(* IEC 61131-3 sources: daoli-st-library/DL_Device (part 29) *)

(* ---- FB_DL_PulseFlowMeter.st ---- *)
(*==============================================================================
 * 组件名称 (Component)  : FB_DL_PulseFlowMeter
 * 所属子库 (Sublibrary) : DL_Device
 * 当前版本 (Version)    : 1.0.0
 * 兼容性   (Platform)   : CODESYS 3.5 / TwinCAT 3 / 汇川 InoProShop / Machine Expert
 *                         仅依赖 Standard.library（TON / R_TRIG），零厂商方言
 * 分类     (Category)   : 设备功能块（Function Block，实现 I_DL_FlowMeter）
 * 功能简述 (Function)   : 脉冲型流量计瞬时流量与累计总量计量。脉冲沿计数 →
 *                         自重触发采样窗频率估计 → K 系数换算 [L/min]；总量
 *                         按脉冲计数法累计（精度优于流量积分法）；低流量截
 *                         止、脉冲丢失超时、频率超量程提示；K 系数防除零。
 *                         滑动窗计数为 Device 层内联实现（依赖方向合规：不
 *                         引 DL_MathData 组件）。
 * 接口实现 (Implements) : I_DL_FlowMeter。接口属性同名成员（eState/fFlowRate/
 *                         fTotal/nPulseCount/bFault/uErrorId）按 R22 以只读
 *                         PROPERTY GET 承载（内部镜像同源），非接口成员
 *                         bTotalNearLimit 保留 VAR_OUTPUT；方法 CmdTotalReset/
 *                         CmdTotalPreset/CmdReset 在本文件尾部落地。
 * 公约遵循 (Convention) : 0.1/R23 周期计量型（无初始化/跟踪同步语义，窗由自
 *                         重触发 TON 驱动），免首扫，无 bInit。
 *                         0.2/R21 bFault 显式排除信息级码；0.5/R7 全部实例主
 *                         体最前部无条件刷新；0.7/R15 故障级锁存仅复位路径清
 *                         码；0.9 全部 REAL/LREAL 输入先做非数自比检测再比
 *                         较，出口默认值在第一条防御 IF 之前赋值。
 *                         0.8 故障码段位 16#0003_xxxx（经 DL_Device
 *                         VERSION.md 码表核对：规格建议信息级 0003_0107/
 *                         0108/0109 已被 FB_DL_VfdGeneric/FB_DL_AnalogValve
 *                         占用，依公约冲突顺延）：
 *                         【故障级】0003_02B0 K 系数非法；
 *                         【信息级】0003_0113 低流量截止激活、0003_0114 脉冲
 *                         丢失超时、0003_0115 窗内频率超量程。
 * 红线自检 (Redline)    : R1 零全局变量表/外部变量引用 ✓｜R2 零物理 IO 地址 ✓
 *                         R3 纯 IEC 61131-3 ✓｜R4 三处除法全部带 ABS(分母)
 *                         >1E-6 防零分支并置码 ✓
 *                         R5 全变量中英双语同行注释 ✓｜R6 状态映像 IF 派生链
 *                         含 ELSE 兜底（无显式 CASE 主状态机，计量型派生映
 *                         像）✓
 *                         R7 四实例（R_TRIG×3/TON×2）主体最前部无条件刷新 ✓
 *                         R8 全常量化 ✓
 * 设计要点 (Key notes)  : ① 瞬时流量 = 窗脉冲数 / 窗秒数 / fKFactor × 60；
 *                         ② 双缓冲：窗运行期脉冲进计数缓冲，窗沿（TON 振荡
 *                           器 Q）整窗交换到读出缓冲，读侧永不撕裂；
 *                         ③ 除零防御三处：fKFactor 非法 → 故障锁存；窗秒数
 *                           由钳位域（100MS~10S）恒非零 + 显式 ABS 防零分支；
 *                           周期法不使用（统一窗法，简化跨平台）；
 *                         ④ 总量按脉冲计数法 fTotal += 窗脉冲数 / fKFactor；
 *                         ⑤ fTotal > 9.0E15 预警（LREAL 整数精度边界）。
 * 偏离留档 (Deviation)  : 依 R11 头注释留档，共 1 条：
 *                         ① 信息级码顺延：规格建议 0003_0107/0108/0109 与既
 *                           有组件冲突，依公约 0.8 顺延为 0003_0113/0114/
 *                           0115（核对结果优先于建议值）。
 * 开源溯源 (Origin)     : 来源标签 tcopen-component / flow-totalizer，T1-1
 *                         OSCAT Basic ◐ 深化旁证（RAW_NOTES_R7 S-6：TcOpen
 *                         流量组件语义域 + OSCAT 流量计窗法计数公开实现思
 *                         想，仅借鉴语义与算法思想；双缓冲、码位与引脚契约
 *                         100% 本库独立设计，clean-room 未复制源码）。
 * 验收向量 (Acceptance) :
 *   V1 已知脉冲序列换算逐拍复算：窗 1S 内 100 脉冲、K=100 → 1.0 L/min；
 *   V2 总量累计与清零：连续 10 窗 @100 脉冲 → fTotal=10.0 L；清零沿 → 0；
 *   V3 低流量截止：fFlowRate < fLowCutoff → 输出置零 + eLowCutoff + 0003_0113；
 *   V4 K 系数非法：fKFactor=0 → 故障锁存 0003_02B0；
 *   V5 脉冲丢失：tPulseTimeout 超时无脉冲 → 流量置零 + 0003_0114；
 *   V6 双缓冲无撕裂推演：窗沿交换拍读侧保持整窗旧值，计数侧从零重启。
 * 修订历史 (Revision)   :
 *   2026-11-15  v1.0.0  首版入库（Round 07 · DL_Device 流量计族实现件）
 *============================================================================*)
FUNCTION_BLOCK FB_DL_PulseFlowMeter IMPLEMENTS I_DL_FlowMeter
VAR_INPUT
    bPulseIn       : BOOL;             // 脉冲输入（Pulse input），R_TRIG 上升沿计数；硬件滤波由输入层保证 / Pulse input, counted on rising edge, HW filtering upstream
    bCmdTotalReset : BOOL;             // 总量清零指令（Total reset command），上升沿生效 / Total reset edge
    fKFactor       : REAL := 100.0;    // 流量计 K 系数（K-factor）[pulses/L]，域 >0，默认 100.0；标定证书值 / K-factor [pulses/L], > 0, calibration value
    tSampleWindow  : TIME := T#1S;     // 频率估计采样窗（Sample window），默认 T#1S，域 100MS~10S 越界钳位；低流量场景增大 / Sample window, clamped 100MS..10S, increase for low flow
    fLowCutoff     : REAL := 0.5;      // 低流量截止阈值（Low-flow cutoff）[L/min]，默认 0.5；低于阈值输出置零 / Low-flow cutoff [L/min], below it the output is zeroed
    tPulseTimeout  : TIME := T#5S;     // 脉冲丢失超时（Pulse timeout），默认 T#5S；运行中窗口超时无脉冲 → 流量置零 + 信息级 / Pulse timeout, no pulse in window zeroes the flow with info
    bReset         : BOOL;             // 上升沿复位故障（Reset edge）/ Rising edge resets fault
END_VAR
VAR_OUTPUT
    bTotalNearLimit : BOOL;            // 总量接近溢出预警（Total near limit），fTotal > 9.0E15 置位（LREAL 整数精度边界）/ Total near LREAL integer-precision boundary
END_VAR
VAR
    _eState        : E_DL_FlowMeterState := E_DL_FlowMeterState.eIdle; // 内部计量状态（Internal metering state），属性只读 / Internal state, read-only via property
    _bFaultLatch   : BOOL;             // 故障锁存标志（Fault latch flag），仅复位路径清除 / Fault latch, cleared only via reset path
    _uErrorIdInt   : UDINT;            // 内部故障级码寄存（Internal fault-level register）/ Internal fault-level register
    _uInfoCode     : UDINT;            // 本拍信息级码（Info code this cycle），瞬时型每拍重算 / Transient info code, recomputed each scan
    _fKFactorEff   : REAL := 100.0;    // 防御后生效 K 系数（Sanitized K-factor）[pulses/L] / Sanitized K-factor
    _fCutoffEff    : REAL := 0.5;      // 防御后生效截止阈值（Sanitized cutoff）[L/min] / Sanitized cutoff
    _tWindowEff    : TIME := T#1S;     // 钳位后生效采样窗（Clamped sample window）/ Clamped sample window
    _nCounting     : UDINT;            // 计数中缓冲（Counting buffer），窗运行期累积 / Counting buffer during the window
    _nLastWin      : UDINT;            // 读出缓冲（Readout buffer），窗沿整窗交换 / Readout buffer swapped at window edge
    _fTotalInt     : LREAL;            // 内部累计总量（Internal totalized volume）[L] / Internal totalized volume [L]
    _fFlowRateInt  : REAL;             // 内部瞬时流量（Internal flow rate）[L/min] / Internal flow rate [L/min]
    _fWinSec       : REAL := 1.0;      // 窗秒数（Window seconds），TIME 显式换算 / Window length in seconds, explicit conversion
    _bHadPulse     : BOOL;             // 曾收到脉冲标志（Ever-pulsed flag），超时判定前提 / Ever-pulsed flag, timeout precondition
    _bPulseLost    : BOOL;             // 脉冲丢失超时激活（Pulse-lost timeout active）/ Pulse-lost timeout active
    _bLowCutoffAct : BOOL;             // 低流量截止激活标志（Low-flow cutoff active flag）/ Low-flow cutoff active flag
    _bPendTotalRst : BOOL;             // 方法总量清零请求（Method total-reset request）/ Method total-reset request
    _bPendPreset   : BOOL;             // 方法总量预置请求（Method total-preset request）/ Method total-preset request
    _fPresetVal    : LREAL;            // 方法预置值（Method preset value）[L] / Method preset value [L]
    _bPendReset    : BOOL;             // 方法复位请求（Method reset request）/ Method reset request
    _fbTrigPulse   : R_TRIG;           // 脉冲上升沿（Pulse rising edge）/ Pulse edge detector
    _fbTrigTotalRst: R_TRIG;           // 引脚总量清零沿（Pin total-reset edge）/ Pin total-reset edge detector
    _fbTrigReset   : R_TRIG;           // 引脚复位沿（Pin reset edge）/ Pin reset edge detector
    _fbTonWindow   : TON;              // 采样窗振荡器（Sample-window oscillator），IN := NOT Q 自重触发 / Sample-window oscillator, self-retriggered
    _fbTonPulseTo  : TON;              // 脉冲丢失超时（Pulse-lost timeout）/ Pulse-lost timeout
END_VAR
VAR CONSTANT
    DL_WIN_MIN     : TIME := T#100MS;  // 采样窗下限（Sample window lower clamp）/ Sample window lower clamp
    DL_WIN_MAX     : TIME := T#10S;    // 采样窗上限（Sample window upper clamp）/ Sample window upper clamp
    DL_PULSE_WIN_MAX : UDINT := 10000; // 单窗脉冲数超量程阈值（Pulses-per-window overrange limit），提示配置 HSC / Per-window pulse overrange, suggests HSC
    DL_TOTAL_LIMIT : LREAL := 9.0E15;  // 总量精度边界预警阈值（Total precision-boundary threshold）[L] / Total precision-boundary threshold [L]
    DL_REAL_EPS    : REAL := 1.0E-6;   // 浮点防零容差（Float divide-guard epsilon）/ Float divide-guard epsilon
END_VAR

METHOD CmdTotalReset : BOOL
VAR_INPUT
END_VAR
IF _bFaultLatch OR (_eState = E_DL_FlowMeterState.eFault) THEN
    CmdTotalReset := FALSE;       // 故障态拒绝（Rejected in fault）
ELSE
    _bPendTotalRst := TRUE;       // 登记清零请求，主体消化（Register reset, consumed by body）
    CmdTotalReset := TRUE;        // 受理成功（Accepted）
END_IF

(*------------------------------------------------------------------------------
 * 方法: CmdTotalPreset —— 总量预置 [L]，非有限值/负值拒绝返回 FALSE。
 *      Method CmdTotalPreset - total preset [L], non-finite or negative rejected.
 *------------------------------------------------------------------------------*)
    END_METHOD

METHOD CmdTotalPreset : BOOL
VAR_INPUT
    fPreset : LREAL; // 预置总量（Preset volume）[L]，域 ≥0 / Preset volume [L], range >= 0
END_VAR
IF _bFaultLatch OR (_eState = E_DL_FlowMeterState.eFault) THEN
    CmdTotalPreset := FALSE;      // 故障态拒绝（Rejected in fault）
ELSIF (fPreset <> fPreset) OR (fPreset < 0.0) THEN
    CmdTotalPreset := FALSE;      // 非数或负值拒绝（Rejected on NaN or negative）
ELSE
    _fPresetVal := fPreset;       // 登记预置值（Register preset value）
    _bPendPreset := TRUE;         // 登记预置请求（Register preset request）
    CmdTotalPreset := TRUE;       // 受理成功（Accepted）
END_IF

(*------------------------------------------------------------------------------
 * 方法: CmdReset —— 复位故障。仅故障态受理（接口方法拒绝语义红线）。
 *      Method CmdReset - reset, accepted only in fault state.
 *------------------------------------------------------------------------------*)
    END_METHOD

METHOD CmdReset : BOOL
VAR_INPUT
END_VAR
IF _bFaultLatch OR (_eState = E_DL_FlowMeterState.eFault) THEN
    _bPendReset := TRUE;          // 登记复位请求（Register reset request）
    CmdReset := TRUE;             // 可复位（Resettable）
ELSE
    CmdReset := FALSE;            // 无故障可复位（Nothing to reset）
END_IF

(*------------------------------------------------------------------------------
 * 属性: eState（GET）—— 当前计量状态只读视图。
 *      Property eState (GET) - read-only metering state view.
 *------------------------------------------------------------------------------*)
    END_METHOD

// ============================================================================
// 段 1｜实例无条件周期刷新（R7/0.5：严禁置于 IF/CASE 分支内）
//      Unconditional per-cycle refresh of all instances (R7/0.5)
// ============================================================================
_fbTrigPulse(CLK    := bPulseIn);
_fbTrigTotalRst(CLK := bCmdTotalReset);
_fbTrigReset(CLK    := bReset);
_fbTonWindow(IN := (NOT _fbTonWindow.Q) AND (NOT _bFaultLatch), PT := _tWindowEff); // 采样窗振荡器（Window oscillator）
_fbTonPulseTo(IN := _bHadPulse AND (NOT _fbTrigPulse.Q) AND (NOT _bFaultLatch), PT := tPulseTimeout); // 脉冲丢失超时（Pulse-lost timeout）

// ============================================================================
// 段 2｜参数防御（0.9：非数自比检测，出口默认值先行）+ 信息级预清零 + 复位
//      Parameter sanitation (0.9) + info preset + reset path
// ============================================================================
_uInfoCode := 0;                  // 信息级瞬时型每拍重算（Transient info recomputed each scan）

IF fKFactor <> fKFactor THEN      // K 系数非数自比检测（K-factor NaN self-compare）
    _bFaultLatch := TRUE;         // K 系数非法锁存（Invalid K-factor latch）
    _uErrorIdInt := 16#0003_02B0; // 0003_02B0 K 系数非法【故障级】/ Invalid K-factor, fault level
ELSIF ABS(fKFactor) <= DL_REAL_EPS THEN
    _bFaultLatch := TRUE;         // K 系数趋零防除零锁存（Near-zero K-factor latch）
    _uErrorIdInt := 16#0003_02B0; // 0003_02B0 K 系数非法【故障级】/ Invalid K-factor, fault level
ELSE
    _fKFactorEff := fKFactor;     // 生效 K 系数镜像（Effective K-factor mirror）
END_IF

IF fLowCutoff <> fLowCutoff THEN  // 截止阈值非数自比（Cutoff NaN self-compare）
    _fCutoffEff := 0.5;           // 回落默认阈值（Fallback default cutoff）
ELSIF fLowCutoff < 0.0 THEN
    _fCutoffEff := 0.0;           // 负值钳零（Negative clamped to zero）
ELSE
    _fCutoffEff := fLowCutoff;    // 生效阈值镜像（Effective cutoff mirror）
END_IF

IF tSampleWindow < DL_WIN_MIN THEN
    _tWindowEff := DL_WIN_MIN;    // 采样窗下限钳位（Window lower clamp）
ELSIF tSampleWindow > DL_WIN_MAX THEN
    _tWindowEff := DL_WIN_MAX;    // 采样窗上限钳位（Window upper clamp）
ELSE
    _tWindowEff := tSampleWindow; // 合法直通（Valid pass-through）
END_IF
_fWinSec := TIME_TO_REAL(_tWindowEff) / 1000.0; // TIME→REAL 换算结果为毫秒数，除 1000 得秒（CODESYS/TwinCAT 口径，舍入意图：整毫秒窗恒精确）/ TIME_TO_REAL yields milliseconds, divide by 1000 for seconds

IF _fbTrigReset.Q OR _bPendReset THEN
    _bPendReset := FALSE;         // 消费方法复位请求（Consume method reset）
    _bFaultLatch := FALSE;        // 故障锁存解除（Fault latch released）
    _uErrorIdInt := 16#0000_0000; // 故障码清零（Fault code cleared）
END_IF

// ============================================================================
// 段 3｜总量清零/预置（引脚沿 + 方法请求）
//      Total reset/preset (pin edge + method request)
// ============================================================================
IF _fbTrigTotalRst.Q OR _bPendTotalRst THEN
    _bPendTotalRst := FALSE;      // 消费方法请求（Consume method request）
    _fTotalInt := 0.0;            // 总量清零（Total cleared）
END_IF
IF _bPendPreset THEN
    _bPendPreset := FALSE;        // 消费方法预置请求（Consume method preset）
    IF _fPresetVal >= 0.0 THEN
        _fTotalInt := _fPresetVal; // 合法预置写入（Valid preset written）
    END_IF                         // 非法预置已被方法拒绝，此处仅兜底（Invalid preset already rejected by method）
END_IF

// ============================================================================
// 段 4｜脉冲计数 + 窗沿双缓冲交换 + 瞬时流量换算（除法全部带防零分支）
//      Pulse counting + double-buffer swap at window edge + flow conversion
// ============================================================================
IF _fbTrigPulse.Q THEN
    _nCounting := _nCounting + 1; // 计数缓冲累加（Counting buffer increment）
    _bHadPulse := TRUE;           // 曾收到脉冲（Ever pulsed）
END_IF

IF _fbTonWindow.Q THEN
    // 窗沿：整窗交换（双缓冲无撕裂：读出缓冲只在窗沿被写一次）
    // Window edge: whole-window swap (readout written once per window, no tearing)
    _nLastWin := _nCounting;      // 读出缓冲接收整窗计数（Readout takes the window count）
    _nCounting := 0;              // 计数缓冲清零重启（Counting buffer restarted）
    IF ABS(_fKFactorEff) > DL_REAL_EPS THEN
        _fTotalInt := _fTotalInt + UDINT_TO_LREAL(_nLastWin) / _fKFactorEff; // 脉冲计数法累计（Count-based totalization, divisor proven non-zero）
    END_IF
END_IF

_fFlowRateInt := 0.0;             // 出口默认值先赋（Default outlet first）
IF ABS(_fWinSec) > DL_REAL_EPS THEN
    IF ABS(_fKFactorEff) > DL_REAL_EPS THEN
        _fFlowRateInt := UDINT_TO_REAL(_nLastWin) / _fWinSec / _fKFactorEff * 60.0; // 窗法换算 [L/min]（Window-method conversion, divisors proven non-zero）
    END_IF
END_IF

// ============================================================================
// 段 5｜诊断与信息级：脉冲丢失 / 频率超量程 / 低流量截止
//      Diagnostics and info codes: pulse lost / overrange / low-flow cutoff
// ============================================================================
_bLowCutoffAct := FALSE;          // 截止激活标志每拍预清零（Cutoff flag preset FALSE）
_bPulseLost := _fbTonPulseTo.Q;   // 脉冲丢失超时激活（Pulse-lost timeout active）
IF _bPulseLost THEN
    _fFlowRateInt := 0.0;         // 超时流量置零（Flow zeroed on timeout）
    _uInfoCode := 16#0003_0114;   // 0003_0114 脉冲丢失超时【信息级】/ Pulse-lost timeout, info level
ELSIF _nLastWin > DL_PULSE_WIN_MAX THEN
    _uInfoCode := 16#0003_0115;   // 0003_0115 窗内频率超量程【信息级】，提示输入层配置 HSC / Per-window overrange, suggest HSC upstream
ELSIF (_fFlowRateInt < _fCutoffEff) AND _bHadPulse AND (NOT _bPulseLost) THEN
    _fFlowRateInt := 0.0;         // 低流量截止输出置零（Low-flow cutoff zeroes output）
    _bLowCutoffAct := TRUE;       // 截止激活标志置位（Cutoff flag asserted）
    _uInfoCode := 16#0003_0113;   // 0003_0113 低流量截止激活【信息级】/ Low-flow cutoff active, info level
END_IF

// ============================================================================
// 段 6｜状态映像（IF 派生链含 ELSE 兜底）+ 输出推导
//      State image (IF derivation chain with ELSE) + output derivation
// ============================================================================
IF _bFaultLatch THEN
    _eState := E_DL_FlowMeterState.eFault;        // 故障映像（Fault image）
ELSIF _bPulseLost OR (NOT _bHadPulse) THEN
    _eState := E_DL_FlowMeterState.eIdle;         // 静默/丢失映像（Idle image）
ELSIF _bLowCutoffAct THEN
    _eState := E_DL_FlowMeterState.eLowCutoff;    // 截止映像（Low-cutoff image）
ELSIF _fFlowRateInt > 0.0 THEN
    _eState := E_DL_FlowMeterState.eFlowOk;       // 正常流量映像（Flow-OK image）
ELSE
    _eState := E_DL_FlowMeterState.eMeasuring;    // 测量中兜底映像（Measuring fallback image）
END_IF

bTotalNearLimit := _fTotalInt > DL_TOTAL_LIMIT; // 总量精度边界预警（Total near precision boundary）

(*------------------------------------------------------------------------------
 * 方法: CmdTotalReset —— 总量清零。故障态拒绝。
 *      Method CmdTotalReset - total reset, rejected in fault.
 *------------------------------------------------------------------------------*)

PROPERTY eState : E_DL_FlowMeterState
eState := _eState;                // 返回内部状态（Return internal state）

(*------------------------------------------------------------------------------
 * 属性: fFlowRate（GET）—— 瞬时流量 [L/min]。
 *      Property fFlowRate (GET) - instantaneous flow rate [L/min].
 *------------------------------------------------------------------------------*)
PROPERTY fFlowRate : REAL
fFlowRate := _fFlowRateInt;       // 返回瞬时流量镜像（Return flow-rate mirror）

(*------------------------------------------------------------------------------
 * 属性: fTotal（GET）—— 累计总量 [L]。
 *      Property fTotal (GET) - totalized volume [L].
 *------------------------------------------------------------------------------*)
PROPERTY fTotal : LREAL
fTotal := _fTotalInt;             // 返回累计总量镜像（Return total mirror）

(*------------------------------------------------------------------------------
 * 属性: nPulseCount（GET）—— 窗口内脉冲计数原始值（读出缓冲）。
 *      Property nPulseCount (GET) - raw pulse count of the last window.
 *------------------------------------------------------------------------------*)
PROPERTY nPulseCount : UDINT
nPulseCount := _nLastWin;         // 返回读出缓冲（Return readout buffer）

(*------------------------------------------------------------------------------
 * 属性: bFault（GET）—— 故障锁存指示（信息级码不置本位，0.2 公约）。
 *      Property bFault (GET) - fault latch indicator, info codes excluded.
 *------------------------------------------------------------------------------*)
PROPERTY bFault : BOOL
bFault := _bFaultLatch OR (_eState = E_DL_FlowMeterState.eFault); // 显式排除信息级派生式（Derived form excluding info codes）

(*------------------------------------------------------------------------------
 * 属性: uErrorId（GET）—— 末次故障码（故障级优先，无故障时透出本拍信息级
 *         码，0.2/0.15 公约）。
 *      Property uErrorId (GET) - last error code (fault priority, info shown otherwise).
 *------------------------------------------------------------------------------*)
PROPERTY uErrorId : UDINT
IF (_uErrorIdInt <> 0) OR (_eState = E_DL_FlowMeterState.eFault) THEN
    uErrorId := _uErrorIdInt;     // 故障级码优先透出（Fault-level priority）
ELSE
    uErrorId := _uInfoCode;       // 无故障时透出本拍信息级码（Transient info code）
END_IF
END_FUNCTION_BLOCK

(* ---- FB_DL_PumpDryRunGuard.st ---- *)
//==============================================================================
// 功能块：FB_DL_PumpDryRunGuard ｜ 中文名称：泵干转保护（双判据 + 防频繁启停）
// 所属子库：DL_Device ｜ 版本：v1.0.1 ｜ 兼容：CODESYS V3.5+ / TwinCAT 3 / 汇川 InoProShop
// 功能描述：泵干转保护三段式——判据（功率 < 干转阈 AND 流量 < 干转阈，
//           双判据同时命中才认定干转，单判据只预警）、去抖（双判据持续
//           tTripDebounce 才跳闸）、防频繁启停（跳闸后 tRestartInh 重启
//           抑制窗 + 运行起步 tLearnWin 启动学习窗内不判干转，避开启动
//           瞬态）。同拍多窗配比约束（R100）：tLearnWin < tTripDebounce
//           < tRestartInh——学习窗必须短于去抖窗，否则启动期永不判干转；
//           重启抑制窗为最长的外层窗。
// 开源溯源 (Origin)：道莅原创实现（参考离心泵干转保护工程惯例（功率/流量双判据） 分类与参数域）
// 单位表：功率[千瓦] / 流量[立方米每小时] / 阈值[同量纲] / 时间[ms]
// 错误码表：16#0003_0188 信息级（干转预警：单判据命中或双判据去抖计窗
//           中，不置 bError）/ 16#0003_0189 信息级（重启抑制窗中：跳闸
//           后防频繁启停计时未满，不置 bError）/ 16#0003_035D 故障级
//           （干转跳闸：双判据 + 去抖窗满，锁存，置 bError）/
//           16#0003_035E 故障级（组态非法：阈值 <= 0、时间窗 <= 0 或
//           任一输入非有限，置 bError）/ 16#0003_035F 故障级兜底（状态机
//           落 ELSE 或非法状态，置 bError）
// 状态机：E_DL_PumpGuardState（六态：eIdle=0 / eRunning=10 / eWarn=20 /
//           eTripped=30 / eInhibit=40 / eFault=99），CASE 含 ELSE 兜底，
//           ELSE 置 035F 并断跳闸输出
// 边界行为：① 组态非法 → 故障态锁存，bReset 复位；② 启动学习窗内
//           （运行反馈上升沿起 tLearnWin）不判干转（启动瞬态豁免）；
//           ③ 跳闸锁存：bTripCmd 保持至 bReset 人工复位（抑制窗满回空闲
//           后仍保持，人工确认复位为唯一清除路径，与④一致）；
//           ④ 使能撤销不自动清跳闸锁存（安全侧：干转须人工确认复位）；
//           ⑤ 单判据命中 → eWarn 预警可观测，判据消失自动回运行态；
//           ⑥ 安全侧 = 故障/空闲路径 bTripCmd := FALSE 且 bValid :=
//           FALSE，跳闸输出只在锁存态保持。
// 修订历史：v1.0.0 2026-11-17 首版（R24 派单 · ROADMAP P1 §452）
//           v1.0.1 2026-11-17 R24 终审修复（R106 第一档，契约不变）：
//           tTripDebounce 默认 3S 与 tLearnWin 默认 5S 自违反头注释
//           R100 配比约束（学习窗 < 去抖窗 < 抑制窗），默认参数出厂即
//           组态非法 035E——默认去抖窗 3S→8S；边界行为③注释与实现
//           漂移同步修正（锁存仅 bReset 清除）。引脚集合与码位不变。
//==============================================================================

(*------------------------------------------------------------------------------
 * 枚举: E_DL_PumpGuardState（归属本功能块，同文件发布，全库唯一定义）
 * 含义: 干转保护相位，每个成员在 CASE 中有且仅有一个标签。
 *-----------------------------------------------------------------------------*)
TYPE E_DL_PumpGuardState :
(
    eIdle     := 0,   // 空闲：泵未运行 / Idle, pump not running
    eRunning  := 10,  // 运行：双判据未命中或学习窗内 / Running, criteria clear or in the learning window
    eWarn     := 20,  // 预警：单判据命中或去抖计窗中 / Warn, one criterion hit or debounce counting
    eTripped  := 30,  // 跳闸：干转锁存，跳闸输出保持 / Tripped, dry-run latched, trip output held
    eInhibit  := 40,  // 抑制：重启抑制窗中（泵已停） / Inhibit, restart window counting, pump stopped
    eFault    := 99   // 故障：组态非法/非法状态 / Fault, illegal config or illegal state
);
END_TYPE

FUNCTION_BLOCK FB_DL_PumpDryRunGuard
VAR_INPUT
    bEnable        : BOOL;                  // 保护使能 [—] / Protection enable
    bReset         : BOOL;                  // 故障复位 [—]，上升沿清跳闸锁存 / Fault reset, rising edge clears the trip latch
    bPumpRunFb     : BOOL;                  // 泵运行反馈 [—] / Pump running feedback
    fMotorPowerKw  : LREAL;                 // 电机功率实测 [千瓦] / Measured motor power [kW]
    fFlowM3h       : LREAL;                 // 流量实测 [立方米每小时] / Measured flow [m3/h]
    fPowerThreshKw : LREAL := 1.0;          // 干转功率阈 [千瓦]，低于此判功率命中，须 > 0 / Dry-run power threshold [kW], must be > 0
    fFlowThreshM3h : LREAL := 0.5;          // 干转流量阈 [立方米每小时]，低于此判流量命中，须 > 0 / Dry-run flow threshold [m3/h], must be > 0
    tTripDebounce  : TIME  := T#8S;         // 双判据去抖窗 [ms]，须 > 0 且 > 学习窗（v1.0.1 默认 3S→8S：原默认 5S 学习窗 > 3S 去抖窗，自违反 R100 配比约束出厂即 035E 故障） / Dual-criteria debounce window [ms], default raised to satisfy learn < debounce < inhibit
    tLearnWin      : TIME  := T#5S;         // 启动学习窗 [ms]，起步瞬态豁免，须 > 0 且 < 去抖窗 / Startup learning window [ms]
    tRestartInh    : TIME  := T#60S;        // 重启抑制窗 [ms]，防频繁启停，须 > 0 且为最长窗 / Restart inhibit window [ms], the longest
END_VAR
VAR_OUTPUT
    bTripCmd       : BOOL;                  // 跳闸指令 [—]（停泵请求，锁存态保持） / Trip command, held while latched
    bRestartBlock  : BOOL;                  // 重启抑制中 [—] / Restart inhibit active
    eState         : E_DL_PumpGuardState;   // 保护相位 [—] / Protection phase
    eErr           : UDINT;                 // 错误码，0 = 无错，码位 16#0003_0188 起信息级、16#0003_035D 起故障级（分带见错误码表） / Error code, 0 = no error, band info/fault per the code table
    bError         : BOOL;                  // 故障级标志，仅故障级错误置位 / Fault-class flag, set only on fault-level codes
    bValid         : BOOL;                  // 输出可用标志 / Outputs usable flag
END_VAR
VAR
    fbDebounce : TON;                       // 双判据去抖计时（每拍无条件刷新）[ms] / Dual-criteria debounce timer, refreshed unconditionally
    fbLearn    : TON;                       // 启动学习窗计时（每拍无条件刷新）[ms] / Startup learning timer, refreshed unconditionally
    fbInhibit  : TON;                       // 重启抑制窗计时（每拍无条件刷新）[ms] / Restart inhibit timer, refreshed unconditionally
    _eState    : E_DL_PumpGuardState := E_DL_PumpGuardState.eIdle; // 当前相位 / Current phase
    _bCfgBad   : BOOL;                      // 组态非法锁存 / Illegal config latch
    _bTripLatch: BOOL;                      // 干转跳闸锁存 / Dry-run trip latch
    _bRunPrev  : BOOL;                      // 运行反馈上拍电平快照（学习窗起步沿） / Previous-scan level of the run feedback
    _bInfoWarn : BOOL;                      // 预警信息当拍标志 / Warn info flag of this scan
    _bInfoInh  : BOOL;                      // 抑制窗信息当拍标志 / Inhibit info flag of this scan
    _bIllegal  : BOOL;                      // 非法状态标志 / Illegal state flag
    _bInit     : BOOL := FALSE;             // 首扫标志，初值 FALSE 取非判定 / First-scan flag, tested negated
END_VAR
VAR CONSTANT
    DL_PDG_INF     : LREAL := 1.7976931348623157E308; // LREAL 幅值上限 / LREAL magnitude ceiling
    DL_PDG_EPS     : LREAL := 1.0E-6;       // 浮点判零容差 [混合] / Float zero tolerance
    DL_PDG_ZERO    : LREAL := 0.0;          // 零值常量，避免裸字面量 [混合] / Zero constant, avoids a bare literal
END_VAR

(*------------------------------------------------------------------------------
 * 段 1｜每拍预置：输出安全侧清零，单拍标志预清零
 *      Outputs cleared fail-safe first, one-shot flags pre-cleared
 *-----------------------------------------------------------------------------*)
bTripCmd      := FALSE;                  // 跳闸指令先清（锁存态在段 6 重置） / Trip command cleared first
bRestartBlock := FALSE;                  // 抑制标志先清 / Inhibit flag cleared first
eErr   := 16#0000_0000;                  // 错误码每拍重算 / Error code recomputed
bError := FALSE;                         // 故障标志每拍重算 / Fault flag recomputed
bValid := FALSE;                         // 可用标志每拍重算 / Usable flag recomputed
_bInfoWarn := FALSE;                     // 预警信息预清零 / Warn info pre-cleared
_bInfoInh  := FALSE;                     // 抑制信息预清零 / Inhibit info pre-cleared
_bIllegal  := FALSE;                     // 非法状态预清零 / Illegal flag pre-cleared

(*------------------------------------------------------------------------------
 * 段 2｜首扫初始化
 *      First-scan initialisation
 *-----------------------------------------------------------------------------*)
IF NOT _bInit THEN
    _eState     := E_DL_PumpGuardState.eIdle; // 相位空闲起步 / Phase starts idle
    _bCfgBad    := FALSE;                  // 组态锁存清零 / Config latch cleared
    _bTripLatch := FALSE;                  // 跳闸锁存清零 / Trip latch cleared
    _bRunPrev   := FALSE;                  // 运行快照清零 / Run snapshot cleared
    _bInit      := TRUE;                   // 首扫只做一次 / The first scan runs once
END_IF

(*------------------------------------------------------------------------------
 * 段 3｜组态防御闸：非有限（R79）+ 阈值/时间窗物理域
 *      Configuration defense gates
 *-----------------------------------------------------------------------------*)
IF (fMotorPowerKw <> fMotorPowerKw) OR (ABS(fMotorPowerKw) > DL_PDG_INF)
   OR (fFlowM3h <> fFlowM3h) OR (ABS(fFlowM3h) > DL_PDG_INF)
   OR (fPowerThreshKw <> fPowerThreshKw) OR (ABS(fPowerThreshKw) > DL_PDG_INF)
   OR (fFlowThreshM3h <> fFlowThreshM3h) OR (ABS(fFlowThreshM3h) > DL_PDG_INF) THEN
    _bCfgBad := TRUE;                      // 非有限归组态非法锁存 / Non-finite folded into the config latch
END_IF
IF (NOT _bCfgBad) AND ((fPowerThreshKw <= DL_PDG_EPS) OR (fFlowThreshM3h <= DL_PDG_EPS)
   OR (tTripDebounce <= T#0MS) OR (tLearnWin <= T#0MS) OR (tRestartInh <= T#0MS)
   OR (tLearnWin >= tTripDebounce) OR (tTripDebounce >= tRestartInh)) THEN
    _bCfgBad := TRUE;                      // 阈值/时间窗非法锁存（含 R100 配比约束：学习窗 < 去抖窗 < 抑制窗） / Threshold and window domains latched with the R100 ratio rule
END_IF

(*------------------------------------------------------------------------------
 * 段 4｜三只计时无条件刷新（R40：CASE 之外每拍必调）
 *      Three timers refreshed unconditionally per R40
 *-----------------------------------------------------------------------------*)
fbDebounce(IN := ((_eState = E_DL_PumpGuardState.eRunning)
                OR (_eState = E_DL_PumpGuardState.eWarn))
           AND (fMotorPowerKw < fPowerThreshKw)
           AND (fFlowM3h < fFlowThreshM3h),
           PT := tTripDebounce);           // 双判据去抖窗（条件含双判据命中） / Debounce window, conditioned on the dual criteria
fbLearn(IN := (_eState = E_DL_PumpGuardState.eRunning)
             OR (_eState = E_DL_PumpGuardState.eWarn),
        PT := tLearnWin);                  // 启动学习窗 / Startup learning window
fbInhibit(IN := (_eState = E_DL_PumpGuardState.eInhibit), PT := tRestartInh); // 重启抑制窗 / Restart inhibit window

(*------------------------------------------------------------------------------
 * 段 5｜相位机（CASE 含 ELSE 兜底；状态改写只出现在分支判据内，R39）
 *      Phase machine with ELSE fallback
 *-----------------------------------------------------------------------------*)
CASE _eState OF

    E_DL_PumpGuardState.eIdle:             // 空闲：运行反馈进运行态
        IF bPumpRunFb AND (NOT _bCfgBad) AND bEnable THEN
            _eState := E_DL_PumpGuardState.eRunning; // 进运行 / To running
        END_IF

    E_DL_PumpGuardState.eRunning:          // 运行：学习窗内豁免；判据命中进预警
        IF (NOT bPumpRunFb) OR (NOT bEnable) OR _bCfgBad THEN
            _eState := E_DL_PumpGuardState.eIdle; // 前置消失回空闲（eWait 类双条件之一） / Precondition gone, back to idle
        ELSIF NOT fbLearn.Q THEN
            _eState := _eState;            // 学习窗内：豁免期不动（显式自持） / Learning window, state held (explicit self-hold)
        ELSIF (fMotorPowerKw < fPowerThreshKw) AND (fFlowM3h < fFlowThreshM3h) THEN
            _bInfoWarn := TRUE;            // 双判据已命中，进预警（拍 N 进入） / Dual criteria hit, to warn
            _eState := E_DL_PumpGuardState.eWarn; // 进预警 / To warn
        ELSIF (fMotorPowerKw < fPowerThreshKw) OR (fFlowM3h < fFlowThreshM3h) THEN
            _bInfoWarn := TRUE;            // 单判据预警（信息级） / Single-criterion warn, info level
        END_IF

    E_DL_PumpGuardState.eWarn:             // 预警：去抖窗满跳闸；判据消失回运行
        IF (NOT bPumpRunFb) OR (NOT bEnable) OR _bCfgBad THEN
            _eState := E_DL_PumpGuardState.eIdle; // 前置消失回空闲 / Precondition gone, back to idle
        ELSIF (fMotorPowerKw >= fPowerThreshKw) AND (fFlowM3h >= fFlowThreshM3h) THEN
            _eState := E_DL_PumpGuardState.eRunning; // 判据消失回运行 / Criteria cleared, back to running
        ELSIF fbDebounce.Q THEN
            _bTripLatch := TRUE;           // 干转跳闸锁存 / Dry-run trip latched
            _eState := E_DL_PumpGuardState.eTripped; // 进跳闸态 / To tripped
        END_IF

    E_DL_PumpGuardState.eTripped:          // 跳闸：输出保持；运行反馈撤销进抑制窗
        IF NOT bPumpRunFb THEN
            _eState := E_DL_PumpGuardState.eInhibit; // 进抑制窗（泵已停） / To inhibit, pump stopped
        END_IF

    E_DL_PumpGuardState.eInhibit:          // 抑制：抑制窗满回空闲（bReset 才清锁存）
        _bInfoInh := TRUE;                 // 抑制窗中（信息级） / Inhibit window active, info
        IF fbInhibit.Q THEN
            _eState := E_DL_PumpGuardState.eIdle; // 抑制窗满回空闲 / Inhibit elapsed, back to idle
        END_IF

    E_DL_PumpGuardState.eFault:            // 故障：复位沿且组态恢复回空闲
        IF bReset AND (NOT _bCfgBad) THEN
            _eState := E_DL_PumpGuardState.eIdle; // 回空闲 / Back to idle
        END_IF

    ELSE                                   // 非法状态兜底（R21：CASE 必带 ELSE）
        _bIllegal := TRUE;                 // 标记非法状态 / Flag the illegal state
        _eState   := E_DL_PumpGuardState.eFault; // 回故障态 / Back to fault
END_CASE
IF bReset THEN
    _bTripLatch := FALSE;                  // 复位清跳闸锁存（人工确认） / Reset clears the trip latch, manual confirmation
END_IF
_bRunPrev := bPumpRunFb;                   // 运行快照推进 / Run snapshot advanced

(*------------------------------------------------------------------------------
 * 段 6｜码位出口与放行（故障级码 3 行内置 bError，R45/R101 配对）
 *      Code outlet and release, fault codes paired with bError
 *-----------------------------------------------------------------------------*)
IF _bIllegal THEN
    eErr   := 16#0003_035F;                // 故障级：状态机兜底 / Fault: state machine fallback
    bError := TRUE;                        // 置故障标志 / Raise the fault flag
ELSIF _bCfgBad THEN
    eErr   := 16#0003_035E;                // 故障级：组态非法 / Fault: illegal configuration
    bError := TRUE;                        // 置故障标志 / Raise the fault flag
ELSIF _bTripLatch THEN
    eErr   := 16#0003_035D;                // 故障级：干转跳闸锁存 / Fault: dry-run trip latched
    bError := TRUE;                        // 置故障标志 / Raise the fault flag
ELSIF _bInfoInh THEN
    eErr := 16#0003_0189;                  // 信息级：重启抑制窗中 / Info: restart inhibit active
ELSIF _bInfoWarn THEN
    eErr := 16#0003_0188;                  // 信息级：干转预警 / Info: dry-run warn
END_IF

bTripCmd := _bTripLatch;                   // 跳闸输出 = 锁存量（不挂单拍标志，R99） / Trip output equals the latch, not a one-shot flag
bRestartBlock := (_eState = E_DL_PumpGuardState.eInhibit); // 抑制中出口 / Inhibit outlet
bValid := (NOT bError) AND bEnable AND (_eState <> E_DL_PumpGuardState.eIdle); // 空闲/故障/未使能输出不可用 / Outputs unusable in idle, fault or disabled
eState := _eState;                         // 相位出口 / Phase outlet
END_FUNCTION_BLOCK

(* ---- FB_DL_PumpDryRunProtect.st ---- *)
(*==============================================================================
 * 组件名称 (Component)  : FB_DL_PumpDryRunProtect
 * 溯源说明 (Provenance) : 道莅 clean-room 防御性实现（Building 泵风机族深化）
 * 所属子库 (Sublibrary) : DL_Device / PumpProtect
 * 当前版本 (Version)    : 1.0.0
 * 兼容性   (Platform)   : CODESYS 3.5 / TwinCAT 3 / 汇川 InoProShop；
 *                         纯 IEC 61131-3（第 3 版），仅用标准库 TON
 * 组件分类 (Category)   : 功能块（FUNCTION_BLOCK）· 泵干转保护
 * 功能一句话 (Summary)  : 运行态功率/流量双判据干转确认 + 确认延时 + 重启闭锁。
 * 边界与安全 (Boundary) : ①仅在运行反馈存在时判定（未运行不判）；
 *                         ②功率与流量任一达到干转特征即计时（双判据并联）；
 *                         ③流量引脚小于 0 表示未接（可选量，仅功率判据）；
 *                         ④空载阈值非正 → 参数非法码；
 *                         ⑤跳闸锁存 + 重启闭锁，需 bReset 且流程恢复才解除。
 * 错误码    : 16#0003_037E 干转确认（延时满足）——故障级（锁存）
 *             16#0003_037F 参数非法（空载阈值非正）——故障级（持续态）
 *             16#0003_0380 重启闭锁激活（跳闸未复位）——故障级（持续态）
 * 码位总账  : 16#0003_037E 用 / 16#0003_037F 用 / 16#0003_0380 用
 * 修改记录  : v1.0.0 R26 初版
 *==============================================================================*)
FUNCTION_BLOCK FB_DL_PumpDryRunProtect
VAR_INPUT
    bPumpRunFb   : BOOL;  // 泵运行反馈 / Pump running feedback
    fMotorPower  : LREAL; // 电机功率 [kW] / Motor power [kW]
    fFlow        : LREAL; // 流量 [m3/h]，小于 0 表示未接 / Flow [m3/h], negative = not wired
    fNoLoadPower : LREAL; // 空载功率阈值 [kW] / No-load power threshold [kW]
    tDryDelay    : TIME;  // 干转确认延时 [ms] / Dry-run confirm delay [ms]
    bReset       : BOOL;  // 复位指令（跳闸后解除闭锁）/ Reset command (clears trip inhibit)
END_VAR
VAR_OUTPUT
    bDryRun        : BOOL; // 干转特征成立（计时中）/ Dry-run signature active (timing)
    bTrip          : BOOL; // 干转跳闸锁存 / Dry-run trip latch
    bRestartInhibit: BOOL; // 重启闭锁（跳闸未复位期间）/ Restart inhibit while latched
    eErr           : UDINT; // 本周期错误码，0=无错 / Error code this cycle, 0 = none
END_VAR
VAR
    tonDry    : TON;   // 干转确认定时器（无条件刷新）/ Dry-run confirm timer
    bPowDry   : BOOL;  // 功率干转特征 / Power dry signature
    bFlowDry  : BOOL;  // 流量干转特征 / Flow dry signature
    bFlowWired: BOOL;  // 流量引脚已接判据 / Flow pin wired predicate
    fPowGuard : LREAL; // 功率守卫副本 / Power guard copy
    fFlowGuard: LREAL; // 流量守卫副本 / Flow guard copy
    bParamOk  : BOOL;  // 参数合法性 / Parameter legality
END_VAR

// ---------- 实时守卫副本 ----------
fPowGuard  := fMotorPower;
fFlowGuard := fFlow;
bFlowWired := fFlowGuard >= 0.0;              // 负值约定为未接 / Negative convention = not wired

// ---------- 参数防御：空载阈值非正或 NaN（持续态，不判定） ----------
bParamOk := (fNoLoadPower > 0.0) AND (fNoLoadPower = fNoLoadPower);
IF NOT bParamOk THEN
    eErr := 16#0003_037F;                     // 参数非法码 / Illegal parameter code
    bDryRun := FALSE;
END_IF

// ---------- 干转双判据：仅运行态判定（未运行不判） ----------
bPowDry  := FALSE;
bFlowDry := FALSE;
IF bPumpRunFb AND bParamOk THEN
    IF (fPowGuard >= 0.0) AND (fPowGuard < fNoLoadPower) THEN
        bPowDry := TRUE;                      // 功率低于空载阈 / Power below no-load threshold
    END_IF
    IF bFlowWired AND (fFlowGuard < 0.01) THEN
        bFlowDry := TRUE;                     // 流量近零 / Flow near zero
    END_IF
END_IF

// ---------- 无条件周期刷新：干转确认定时器 ----------
tonDry(IN := bPowDry OR bFlowDry, PT := tDryDelay);
bDryRun := tonDry.IN;                         // 计时中特征输出 / Signature while timing

// ---------- 跳闸锁存与重启闭锁 ----------
IF tonDry.Q THEN
    bTrip := TRUE;                            // 延时满足跳闸锁存 / Delay met, trip latch
    eErr  := 16#0003_037E;                    // 干转确认码 / Dry-run confirm code
END_IF

IF bTrip THEN
    bRestartInhibit := TRUE;                  // 闭锁激活 / Inhibit active
    eErr := 16#0003_0380;                     // 重启闭锁码（跳闸确认码 037E 已在确认拍报出）/ Inhibit code, trip code raised at confirm scan
    IF bReset THEN
        bTrip           := FALSE;             // 复位解除锁存 / Reset clears latch
        bRestartInhibit := FALSE;             // 闭锁解除 / Inhibit cleared
        eErr            := 0;                 // 复位同拍清码 / Code cleared on reset
    END_IF
ELSE
    bRestartInhibit := FALSE;                 // 无锁存无闭锁 / No latch, no inhibit
END_IF

END_FUNCTION_BLOCK

(* ---- FB_DL_PumpPrimingWatch.st ---- *)
(*
    FB_DL_PumpPrimingWatch —— 离心泵灌泵期监视（充水确认窗 + 起立判据 + 干转前预警）
    ------------------------------------------------------------------
    组件名称  : FB_DL_PumpPrimingWatch
    分类      : DL_Device / PumpHealth
    前缀      : FB_DL_
    版本      : 1.0.0
    溯源      : 借鉴点 —— 内部台账 T2-2 行「命令 - 监视 - 判定」三段分层骨架
                （R11 / R13 先例，self 判据）。
                本件只借**骨架**，灌泵窗口 / 双判据 / 码位 100% 自有。
                clean-room 声明 —— 零代码行复制；定时与沿检测仅用 IEC 61131-3
                标准库 TON / R_TRIG。
                许可证 —— 本件 MIT；来源标签 t2-2-lbp 为闭源内部台账，
                按最严口径零代码行接触。
    平台      : 纯 IEC 61131-3，CODESYS 3.5 / TwinCAT 3 / InoProShop / Machine Expert 通用
    作者      : 道莅代码库 · PLC编程专家（R71 构建轮 · 批 2 · 序号 8）
    ------------------------------------------------------------------
    功能说明  : 灌泵期（启动前充水确认）监视顺控：
                eIdle 待机 →（bStartCmd 上升沿）ePriming 灌泵确认窗计时
                →（流量 ∧ 压力双判据同拍持续 tConfirm）ePrimed 灌泵完成放行
                →（命令撤销）eIdle；窗满仍无起立 → ePrimeFail 失败相 +
                锁存码（干转前预警，锁存待复位）。
                双窗设计（R41 / R42 口径）：
                _tonWin 灌泵总窗（PT = tPrimeWin，IN = 相为 ePriming），
                _tonCfm 起立判据驻留确认（PT = tConfirm，IN = 相为 ePriming
                且流量 ∧ 压力本拍实时复验成立）——两实例每周期无条件调用，
                IN 为显式条件，选窗不依赖可跳过分支。
                窗满迁移判据（R41 同拍竞态收敛）：失败 = 窗满 ∧ 反馈**仍**
                无效（窗满拍复验一次）；反馈迟到但在窗满拍有效 → 不判失败，
                由 _tonCfm 驻留确认路径继续收敛至 ePrimed（驻留上限
                tConfirm 有界，不会无限延窗）。
                起立判据「先判后信」（R42）：bFlowOK / bPressOK 为本拍复验的
                实时反馈，沿上不锁存旧反馈。
                失败锁存语义：ePrimeFail 相锁存（37C1），bReset 上升沿唯一
                解除回 eIdle —— 干转前预警属安全结论，不允许命令撤销顺手
                清除（R303 失能不清锁存同口径）。
    错误码    : 16#0002_37C0 组态非法（tPrimeWin / tConfirm 非正，或
                            tConfirm >= tPrimeWin 配比吞没失败判据），锁存
                            —— 故障级
                16#0002_37C1 灌泵窗满且起立判据仍无效（干转前预警），锁存
                            —— 故障级
                16#0002_37C2 非法相枚举（CASE ELSE 兜底），锁存 —— 故障级
    码位总账  : 37C0 / 37C1 / 37C2 用（均故障级，本件无信息级码）
    状态机    : ENUM E_DL_PpwPhase 五态，CASE 全覆盖 + ELSE 兜底（锁存 37C2
                回 eFault）。迁移表见功能说明；bReset 上升沿：解锁存（含
                ePrimeFail）→ eIdle（唯一可到达的解除边，R188）。
    边界与披露: 一 组态判据逐项点名（R272）：tPrimeWin <= T#0S 拦截；
                   tConfirm < T#0S 拦截（TIME 非负语义下的防御复检）；
                   **同拍双窗配比约束（R100）：tConfirm >= tPrimeWin 拦截** ——
                   确认驻留窗大于等于总窗时，失败判据（窗满 ∧ 反馈无效）
                   永不成立，干转预警静默失效，属组态级禁止；
                二 布尔反馈输入（bFlowOK / bPressOK / bStartCmd）无非有限面，
                   不设数值闸；反馈真值即判据源，无换算无死区（无魔法数）；
                三 失能（bEn = FALSE）语义写死（R303）：bPriming / bPrimed /
                   bPrimeFail 输出全清零、bError 清零、码清零、状态回 eIdle，
                   但 _bFault 锁存位**不被失能清除**（失能是操作态，不是
                   复位），必须 bReset 上升沿才解除 —— 两者语义分离；
                四 定时器 _tonWin / _tonCfm 无论失能 / 故障 / 正常均在段 7
                   无条件调用，IN 为段 6 计算出的显式条件；
                五 ePrimed 相命令撤销即回 eIdle（电平判定，非沿 —— 命令
                   保持则持续放行，命令撤销即收回放行资格，名实一致）；
                六 零全局变量、零 VAR_EXTERNAL、零物理地址、零数组下标、
                   无除法、无浮点量。
    分工声明  : FB_DL_PumpDryRunProtect（DL_Device，运行期干转保护）、
                FB_DL_PumpCavitationGuard（DL_Device，运行期汽蚀防护）、
                FB_DL_PumpAlternationLead（DL_Process，多泵轮值）——本件专管
                **灌泵期**（启动前充水确认），运行期判据归既有三件，
                四者互引分工边界，不互代。
    修订记录  : 2026-11-22 v1.0.0 首次入库（R71 构建轮 · 批 2 · 序号 8）
*)
TYPE E_DL_PpwPhase :
(
    eIdle      := 0,   (* 待机，等启泵命令沿 / idle, waiting for a start command edge *)
    ePriming   := 10,  (* 灌泵确认窗相（双窗计时 + 起立判据监视）/ the priming phase, the dual window timing plus the primed criteria watch *)
    ePrimed    := 20,  (* 灌泵完成相（放行，命令撤销即回待机）/ the primed phase, released, back to idle on command withdrawal *)
    ePrimeFail := 30,  (* 灌泵失败相（窗满无起立，锁存待复位）/ the prime fail phase, the window full without priming, latched for a reset *)
    eFault     := 40   (* 故障相（非法枚举兜底锁存）/ the fault phase, the illegal enumeration guard latch *)
);
END_TYPE

FUNCTION_BLOCK FB_DL_PumpPrimingWatch
VAR_INPUT
    bEn       : BOOL := TRUE;              (* 使能，[标志]，FALSE 时出口清零且状态回待机（R303）/ the enable, FALSE clears the outlets and returns to idle *)
    bReset    : BOOL := FALSE;             (* 故障 / 失败复位（上升沿有效），[标志] / the reset, rising edge effective, the only release *)
    bStartCmd : BOOL := FALSE;             (* 启泵命令（上升沿启动 / 电平保持放行），[标志] / the pump start command *)
    bFlowOK   : BOOL := FALSE;             (* 流量起立反馈（本拍实时复验），[标志] / the flow established feedback, verified live this scan *)
    bPressOK  : BOOL := FALSE;             (* 压力起立反馈（本拍实时复验），[标志] / the pressure established feedback, verified live this scan *)
    tPrimeWin : TIME := T#10S;             (* 灌泵确认总窗，[ms]，须 > T#0S / the priming window *)
    tConfirm  : TIME := T#2S;              (* 起立判据驻留确认时长，[ms]，须 < tPrimeWin（配比约束）/ the criteria hold duration, must be under tPrimeWin *)
END_VAR
VAR_OUTPUT
    eState    : E_DL_PpwPhase := E_DL_PpwPhase.eIdle; (* 相状态出口，[相] / the phase outlet *)
    bPriming  : BOOL;                      (* 灌泵进行中（确认窗计时相），[标志] / the priming in progress flag *)
    bPrimed   : BOOL;                      (* 灌泵完成放行，[标志] / the primed release flag *)
    bPrimeFail: BOOL;                      (* 灌泵失败（干转前预警，锁存），[标志] / the prime fail flag, latched *)
    bError    : BOOL;                      (* 故障标志，锁存故障时为 TRUE / the fault flag, raised while latched *)
    nErrCode  : UDINT;                     (* 错误码，0 = 正常，锁存回放 / the error id, 0 = ok, replayed from the latch *)
END_VAR
VAR
    _rtStart    : R_TRIG;                  (* 启泵命令上升沿实例（无条件调用）/ the start command rising edge instance *)
    _rtReset    : R_TRIG;                  (* 复位上升沿实例（无条件调用）/ the reset rising edge instance *)
    _tonWin     : TON;                     (* 灌泵总窗实例（无条件调用）/ the priming window timer *)
    _tonCfm     : TON;                     (* 起立判据驻留确认实例（无条件调用）/ the criteria hold confirmation timer *)
    _ePhase     : E_DL_PpwPhase := E_DL_PpwPhase.eIdle; (* 相状态寄存器 / the internal phase register *)
    _bFault     : BOOL;                    (* 故障锁存位（含灌泵失败锁存），仅 bReset 上升沿解除 / the latched fault bit, including the prime fail latch *)
    _nCodeLatch : UDINT;                   (* 锁存成因码，故障期回放 / the latched cause code, replayed *)
    _bCfgBad    : BOOL;                    (* 组态非法标志（逐拍重算）/ the configuration fault flag *)
    _bCriteria  : BOOL;                    (* 起立判据本拍复验值（流量 ∧ 压力）/ the primed criteria verified this scan *)
END_VAR

// 段 1｜出口预置（R256 统一出口预置）/ segment 1, preset every outlet
eState    := _ePhase;                     // 相出口先镜像寄存器 / mirror the phase register first
bPriming  := FALSE;                       // 灌泵进行中预清零 / preset the priming flag false
bPrimed   := FALSE;                       // 放行预清零 / preset the primed flag false
bPrimeFail:= FALSE;                       // 失败预清零 / preset the fail flag false
bError    := FALSE;                       // 故障标志预清零 / preset the error flag false
nErrCode  := 0;                           // 错误码预置无错 / preset the code to zero
_bCriteria:= FALSE;                       // 起立判据预清零 / preset the criteria false

// 段 2｜沿检测实例无条件调用（规则 ⑦）/ segment 2, the edge instances, called unconditionally
_rtStart(CLK := bStartCmd);               // 启泵沿，每周期无条件刷新 / the start edge, refreshed every scan
_rtReset(CLK := bReset);                  // 复位沿，每周期无条件刷新 / the reset edge, refreshed every scan

// 段 3｜锁存解除：仅 bReset 上升沿，锁存码同步清零（唯一解除边，R188）/ segment 3, the only latch release edge
IF _rtReset.Q THEN                        // 复位上升沿 / the reset rising edge
    _bFault     := FALSE;                 // 解除故障锁存（含灌泵失败）/ release the fault latch, including the prime fail
    _nCodeLatch := 0;                     // 清锁存码（可到达的清除边）/ clear the latched code, a reachable clearing edge
    _ePhase     := E_DL_PpwPhase.eIdle;   // 回待机相（安全相）/ back to the safe idle phase
END_IF

// 段 4｜组态守卫（边界一逐项点名 + 双窗配比约束，R272 / R100）/ segment 4, the configuration guard
_bCfgBad := (tPrimeWin <= T#0S)           // 总窗非正 / a non positive window
         OR (tConfirm < T#0S)             // 驻留为负（TIME 非负语义下的防御复检）/ a negative hold duration
         OR (tConfirm >= tPrimeWin);      // 配比约束：驻留吞没总窗 → 失败判据永不成立（干转预警静默失效）/ the hold swallows the window, the fail verdict unreachable

// 段 5｜首次成因锁存（故障期不重推断，回放锁存码，R189）/ segment 5, the first-cause latch
IF NOT _bFault THEN                       // 未锁存才登记成因 / a cause is registered only while not latched
    IF _bCfgBad THEN                      // 组态非法（根因）/ the configuration, the root cause
        _bFault     := TRUE;              // 置锁存 / latch it
        _nCodeLatch := 16#0002_37C0;      // 故障级：组态非法 / fault level: an illegal configuration
        _ePhase     := E_DL_PpwPhase.eFault; // 迁入故障相 / enter the fault phase
    END_IF
END_IF

// 段 6｜起立判据本拍复验（R42 先判后信，显式条件供定时器与状态机共用）/ segment 6, the criteria verified this scan
_bCriteria := bFlowOK AND bPressOK;       // 流量 ∧ 压力双判据同拍成立 / the flow and the pressure both hold this scan

// 段 7｜双定时器无条件周期调用（规则 ⑦，IN 为显式条件）/ segment 7, the dual timers, called unconditionally
_tonWin(IN := (_ePhase = E_DL_PpwPhase.ePriming), PT := tPrimeWin);  // 灌泵总窗计时 / the priming window timer
_tonCfm(IN := ((_ePhase = E_DL_PpwPhase.ePriming) AND _bCriteria), PT := tConfirm); // 驻留确认计时 / the hold confirmation timer

// 段 8｜失能相输出回夹（R57 + R303，先于状态机执行）/ segment 8, the disable phase output clamping
IF (NOT bEn) AND (NOT _bFault) THEN       // 失能且无锁存故障（操作态不发码）/ disabled without a latched fault
    _ePhase := E_DL_PpwPhase.eIdle;       // 状态回待机 / back to idle
END_IF                                    // 输出清零由段 1 预置 + 状态机仅在运行许可时执行共同保证

// 段 9｜相状态机（ENUM + CASE + ELSE 兜底，仅运行许可时执行）/ segment 9, the phase machine, run permit only
IF bEn AND NOT _bFault THEN               // 运行许可成立 / the run permit holds
CASE _ePhase OF
    E_DL_PpwPhase.eIdle:                  // 待机相 / the idle phase
        IF _rtStart.Q THEN                // 启泵命令上升沿 / a start command edge
            _ePhase := E_DL_PpwPhase.ePriming; // 进入灌泵确认窗相 / enter the priming phase
        END_IF
    E_DL_PpwPhase.ePriming:               // 灌泵确认窗相 / the priming phase
        IF _tonCfm.Q THEN                 // 起立判据驻留确认完成（双判据持续 tConfirm）/ the criteria hold confirmed
            _ePhase := E_DL_PpwPhase.ePrimed; // 进入灌泵完成相 / enter the primed phase
        ELSIF _tonWin.Q AND (NOT _bCriteria) THEN // 窗满拍复验一次：反馈仍无效才判失败（R41 同拍竞态收敛）/ the window full and the feedback still invalid
            _bFault     := TRUE;          // 锁存故障（干转前预警）/ latch the fault
            _nCodeLatch := 16#0002_37C1;  // 故障级：窗满无起立 / fault level: the window full without priming
            _ePhase     := E_DL_PpwPhase.ePrimeFail; // 迁入失败相（锁存待复位）/ enter the prime fail phase
        END_IF                            // 窗满但反馈已有效 → 不判失败，驻留路径继续收敛（有界 tConfirm）
    E_DL_PpwPhase.ePrimed:                // 灌泵完成相（放行）/ the primed phase
        IF NOT bStartCmd THEN             // 命令撤销（电平判定，边界五）/ the command withdrawn, a level verdict
            _ePhase := E_DL_PpwPhase.eIdle; // 回待机（放行资格随预置收回）/ back to idle, the release withdrawn by the preset
        END_IF
    E_DL_PpwPhase.ePrimeFail:             // 灌泵失败相（锁存保持）/ the prime fail phase, latched
        bError   := TRUE;                 // 故障标志置位 / raise the fault flag
        nErrCode := _nCodeLatch;          // 回放锁存码（不按当下输入重推断）/ replay the latched code
    E_DL_PpwPhase.eFault:                 // 故障相（锁存保持）/ the fault phase, latched
        bError   := TRUE;                 // 故障标志置位 / raise the fault flag
        nErrCode := _nCodeLatch;          // 回放锁存码 / replay the latched code
    ELSE                                  // 非法枚举兜底（回安全相 + 置码，规则 ⑥）/ the illegal enumeration guard
        _bFault     := TRUE;              // 置锁存 / latch it
        _nCodeLatch := 16#0002_37C2;      // 故障级：非法相枚举 / fault level: an illegal phase value
        _ePhase     := E_DL_PpwPhase.eFault; // 回安全相（故障相）/ force the safe fault phase
        bError      := TRUE;              // 故障标志置位（禁静默）/ raise the flag
        nErrCode    := _nCodeLatch;       // 回放锁存码 / replay the latched code
END_CASE
END_IF

// 段 10｜出口映射（名实双出口同源，单点写入，R191）/ segment 10, the outlet mapping
bPriming   := (_ePhase = E_DL_PpwPhase.ePriming); // 灌泵进行中出口与相寄存器同源 / the priming outlet shares the register
bPrimed    := (_ePhase = E_DL_PpwPhase.ePrimed);    // 放行出口与相寄存器同源 / the primed outlet shares the register
bPrimeFail := (_ePhase = E_DL_PpwPhase.ePrimeFail); // 失败出口与相寄存器同源 / the fail outlet shares the register
eState     := _ePhase;                    // 相出口 = 寄存器（段 9 之后不再触碰）/ the phase outlet, not touched after segment 9
IF _bFault THEN                           // 锁存故障相出口补充 / the latched fault supplement
    bError   := TRUE;                     // 故障标志 / the fault flag
    nErrCode := _nCodeLatch;              // 回放锁存码 / replay the latched code
END_IF
END_FUNCTION_BLOCK

(* ---- FB_DL_QuenchTankAgitatorCtrl.st ---- *)
(*
  Component : FB_DL_QuenchTankAgitatorCtrl
  Category  : DL_Device
  Type      : FB
  Complexity: C2
  VERSION   : v1.0.0
  功能      : 淬火槽搅拌器分级投运控制：按油温分三级递增投运，超温持续超时联锁停泵并锁存，R_TRIG 捕捉升入二级的上升沿上报信息码。
  开源溯源  : 道莅原创 clean-room 自研（无外部代码引用）｜License: MIT
  边界条件  : ① 三级温度阈值必须严格递增且低于联锁温度，否则判组态非法并锁存故障；
              ② 超温联锁为持续型判据（延时确认），复位后若温度仍超限将立即重新锁存；
              ③ 泵输出为互锁递进：N 级投运时前 N 台全部运行，高液位/超温时全部切除。
*)
FUNCTION_BLOCK FB_DL_QuenchTankAgitatorCtrl
VAR_INPUT
    bEnable    : BOOL;   (* 使能电平 [-] Enable level *)
    bReset     : BOOL;   (* 复位上升沿，清联锁锁存 [-] Reset edge *)
    fOilTempC  : REAL;   (* 油槽实测油温 [°C] Measured oil temperature *)
    fStage1C   : REAL;   (* 一级投运温度 [°C] Stage 1 start temperature *)
    fStage2C   : REAL;   (* 二级投运温度 [°C] Stage 2 start temperature *)
    fStage3C   : REAL;   (* 三级投运温度 [°C] Stage 3 start temperature *)
    fTripC     : REAL;   (* 超温联锁温度 [°C] Over-temperature trip limit *)
    tTripDelay : TIME;   (* 超温确认延时 [ms] Trip confirmation delay *)
END_VAR
VAR_OUTPUT
    bPump1  : BOOL;    (* 一级搅拌泵输出 [-] Agitator pump 1 output *)
    bPump2  : BOOL;    (* 二级搅拌泵输出 [-] Agitator pump 2 output *)
    bPump3  : BOOL;    (* 三级搅拌泵输出 [-] Agitator pump 3 output *)
    nStage  : INT;     (* 当前投运级数 0~3 [-] Active stage count *)
    bTrip   : BOOL;    (* 超温联锁锁存标志 [-] Trip latch flag *)
    bError  : BOOL;    (* 故障锁存标志 [-] Fault latch flag *)
    uErrId  : UDINT;   (* 事件码，0 = 无事件 [-] Event code *)
END_VAR
VAR
    rtReset    : R_TRIG;  (* 复位沿实例，每拍无条件刷新 / Reset edge *)
    rtStage2   : R_TRIG;  (* 升入二级上升沿实例 / Stage-2 rising edge *)
    tonTrip    : TON;     (* 超温确认计时（独立实例） / Trip confirmation timer *)
    _bTrip     : BOOL;    (* 联锁锁存位（锁存量） / Latched trip bit *)
    _bFault    : BOOL;    (* 故障锁存位（锁存量） / Latched fault bit *)
    _uFault    : UDINT;   (* 故障码锁存（锁存量） / Latched fault code *)
    _bS2Rise   : BOOL;    (* 二级上升沿单拍位 [-] Stage-2 rise one-shot *)
    _bCfgBad   : BOOL;    (* 组态非法当拍量 [-] Config illegal flag *)
    _bNonFin   : BOOL;    (* 输入非有限当拍量 [-] Non-finite input flag *)
END_VAR
VAR CONSTANT
    DL_EPS : REAL := 1.0E-9;   (* 浮点比较容差 [无量纲] Float compare tolerance *)
END_VAR

(* —— 段 1｜每拍量预清零（锁存量 _bTrip/_bFault/_uFault 不入清单） —— *)
uErrId := 16#0000_0000;
_bS2Rise := FALSE;
_bCfgBad := FALSE;
_bNonFin := FALSE;
nStage := 0;

(* —— 段 2｜输入非有限拦截 —— *)
IF (fOilTempC <> fOilTempC) OR ((fOilTempC - fOilTempC) <> 0.0) THEN
    _bNonFin := TRUE;
END_IF

(* —— 段 3｜组态闸：三级阈值严格递增且低于联锁温度，全部参与判据的引脚逐个覆盖 —— *)
IF (fStage1C >= fStage2C) OR (fStage2C >= fStage3C) OR (fStage3C >= fTripC) THEN
    _bCfgBad := TRUE;
END_IF

(* —— 段 4｜温度分级判定（无 NaN 时执行；分组阶梯，不插值） —— *)
IF (NOT _bNonFin) AND (NOT _bCfgBad) THEN
    IF fOilTempC > (fStage3C + DL_EPS) THEN
        nStage := 3;                     (* 三级投运 [-] / Stage 3 *)
    ELSIF fOilTempC > (fStage2C + DL_EPS) THEN
        nStage := 2;                     (* 二级投运 [-] / Stage 2 *)
    ELSIF fOilTempC > (fStage1C + DL_EPS) THEN
        nStage := 1;                     (* 一级投运 [-] / Stage 1 *)
    ELSE
        nStage := 0;                     (* 全部停运 [-] / All stopped *)
    END_IF
END_IF

(* —— 段 5｜沿与定时器每拍无条件刷新（禁置于 IF/CASE 内，使能挂 IN 引脚） —— *)
rtReset (CLK := bReset);
rtStage2(CLK := (nStage >= 2));
tonTrip (IN := _bNonFin OR ((fOilTempC >= fTripC) AND bEnable), PT := tTripDelay);

IF rtStage2.Q THEN
    _bS2Rise := TRUE;                    (* 升入二级上升沿捕获，出口单拍映射 *)
END_IF

(* —— 段 6｜复位沿：联锁与故障一次性清干净（唯一解除路径，恒可达） —— *)
IF rtReset.Q THEN
    _bTrip := FALSE;
    _bFault := FALSE;
    _uFault := 16#0000_0000;
END_IF

(* —— 段 7｜超温联锁：延时确认后锁存，锁存量不当拍按输入重算 —— *)
IF (NOT _bTrip) AND tonTrip.Q THEN
    _bTrip := TRUE;
END_IF
IF (NOT _bFault) AND _bCfgBad THEN
    _bFault := TRUE;
    _uFault := 16#0021_0001;             (* 故障级：温度阈值组态非法 / Bad threshold config *)
END_IF
IF (NOT _bFault) AND _bNonFin THEN
    _bFault := TRUE;
    _uFault := 16#0021_0002;             (* 故障级：油温反馈非有限 / Non-finite temperature *)
END_IF

(* —— 段 8｜输出侧：使能、联锁、故障三者全通过才允许投运 —— *)
IF bEnable AND (NOT _bTrip) AND (NOT _bFault) THEN
    bPump1 := nStage >= 1;               (* 一级泵 [-] / Pump 1 *)
    bPump2 := nStage >= 2;               (* 二级泵 [-] / Pump 2 *)
    bPump3 := nStage >= 3;               (* 三级泵 [-] / Pump 3 *)
ELSE
    bPump1 := FALSE;                     (* 安全侧切除 [-] / Cut off to safe side *)
    bPump2 := FALSE;
    bPump3 := FALSE;
END_IF

(* —— 段 9｜出口单点映射（锁存码回放 + 信息码单拍） —— *)
bTrip := _bTrip;
bError := _bFault;
IF _bFault AND (_uFault <> 16#0000_0000) THEN
    uErrId := _uFault;                   (* 故障码锁存回放 / Latched fault replay *)
ELSIF _bS2Rise THEN
    uErrId := 16#0021_0101;              (* 信息级：升入二级搅拌投运沿 / Stage-2 rise info *)
END_IF
END_FUNCTION_BLOCK

(* ---- FB_DL_RackDiagSummary.st ---- *)
// =====================================================================
// FB_DL_RackDiagSummary.st
// 机架诊断汇总与首出定位（板级状态字聚合 + 首出三律 + 诊断风暴提示）
// Rack diagnostics aggregation with first-out location and storm hint
// 所属子库: DL_Device    版本: v1.0.0    兼容: CODESYS V3.5+ / TwinCAT 3 / 汇川 InoProShop
// 码位: 16#0003_03ED ~ 16#0003_03F1 (本件独占 5 槽, 勿复用)
// 溯源: 道莅 clean-room 防御性实现
//       来源组标签: diagnostics, axioline, first-out, rack
// 修改记录: R30 初版 (ROUND_PLAN_R30 序 5)
// 注: 板级诊断状态字经输入引脚注入, 零外部系统变量依赖, 与库内端口诊断
//     聚合件和单板诊断锁存件的契约字段语义一一对应, 同名位语义不复定义
// =====================================================================
FUNCTION_BLOCK FB_DL_RackDiagSummary
VAR_INPUT
    auBoardStat : ARRAY[1..8] OF WORD;  // 各板卡诊断状态字注入, 非 0 即该板存在故障 / Per-board status word injected, nonzero = fault
    bReset      : BOOL  := FALSE;       // 首出复位命令 / First-out reset command
END_VAR
VAR_OUTPUT
    uwFaultMask : WORD   := 0;          // 板级故障掩码, 位 0..7 对应板 1..8 / Board fault mask, bit0..7 = board 1..8
    uFirstBoard : USINT  := 0;          // 首出板号 1~8, 0 = 无 / First-out board 1..8, 0 = none
    uFirstCode  : UDINT  := 0;          // 首出板状态字快照回放 / First-out board status snapshot replay
    bStorm      : BOOL   := FALSE;      // 诊断风暴单拍标志, 不锁存不置故障级 / Storm single-cycle flag, info only
    eErr        : UDINT  := 16#0003_03ED;  // 错误码 / Error code
END_VAR
VAR
    rtrReset    : R_TRIG;               // 复位上升沿检测, 每拍无条件刷新 / Reset edge, refreshed every cycle
    uwPrevMask  : WORD   := 0;          // 上拍故障掩码快照 / Previous cycle mask snapshot
    uNewCnt     : USINT  := 0;          // 本拍新故障板数 / New fault board count this cycle
    wBit        : WORD   := 0;          // 位测试掩码 / Bit test mask
    bAllFault   : BOOL   := FALSE;      // 全板故障标记 / All-boards-fault flag
    uZi         : INT    := 1;          // 1..8 数组下标 / Array subscript 1..8
END_VAR

// ---------------------------------------------------------------------
// 代码位表（本件独占, 勿复用）:
//   16#0003_03ED 信息 全部板卡无故障
//   16#0003_03EE 信息 诊断风暴提示（单拍新故障板数不小于 4, 仅提示, 不进入故障级）
//   16#0003_03EF 故障 存在板卡故障（掩码非零）, 解除式 = 对应板状态字归零
//   16#0003_03F0 故障 首出锁定有效（板号与状态字快照持续回放）,
//                解除式 = bReset 上升沿 且 首出板故障位已消失
//   16#0003_03F1 故障 全部 8 块板卡故障（整架失效）
// ---------------------------------------------------------------------

// ---- 逐板故障判与掩码聚合 / Per-board fault judge and mask aggregation ----
uwFaultMask := 0;                   // 掩码复位 / Reset mask
FOR uZi := 1 TO 8 DO
    IF auBoardStat[uZi] <> 0 THEN
        uwFaultMask := uwFaultMask OR SHL(WORD#1, uZi - 1);     // 移位量 0..7 小于字宽, 合规 / Shift within word width
    END_IF
END_FOR

// ---- 本拍新故障板数差分（与上拍掩码比对）/ New fault count vs previous mask ----
uNewCnt := 0;                       // 新故障计数复位 / Reset new fault count
FOR uZi := 1 TO 8 DO
    wBit := SHL(WORD#1, uZi - 1);   // 当前板位掩码 / Current board bit mask
    IF (uwFaultMask AND wBit) <> 0 THEN
        IF (uwPrevMask AND wBit) = 0 THEN
            uNewCnt := uNewCnt + 1; // 本拍新出现故障的板 / Newly faulted board this cycle
        END_IF
    END_IF
END_FOR
bStorm := uNewCnt >= 4;             // 单拍新故障板数达 4 判风暴, 单拍标志当拍自清 / Storm if 4+ new per cycle
uwPrevMask := uwFaultMask;          // 快照更新供下拍差分 / Snapshot for next cycle

// ---- 复位沿实例无条件刷新 / Unconditional reset edge refresh ----
rtrReset(CLK := bReset);

// ---- 首出三律: 未锁存才仲裁, 同拍取最小板号, 解除在仲裁后 / First-out three laws ----
IF uFirstBoard = 0 THEN
    FOR uZi := 1 TO 8 DO
        IF (uFirstBoard = 0) AND ((uwFaultMask AND SHL(WORD#1, uZi - 1)) <> 0) THEN
            uFirstBoard := INT_TO_USINT(uZi);                   // 升序扫描取最小板号 / Ascending scan picks min board
            uFirstCode  := WORD_TO_UDINT(auBoardStat[uZi]);     // 锁存首出板状态字快照 / Latch status snapshot
        END_IF
    END_FOR
END_IF
// 解除式: bReset 上升沿 且 首出板故障位已消失 / Release: reset edge AND first-out fault bit gone
IF rtrReset.Q AND (uFirstBoard <> 0)
   AND ((uwFaultMask AND SHL(WORD#1, uFirstBoard - 1)) = 0) THEN
    uFirstBoard := 0;               // 释放首出板号 / Release first-out board
    uFirstCode  := 0;               // 清状态字快照 / Clear snapshot
END_IF

// ---- 全板故障判 / All-boards-fault judge ----
bAllFault := (uwFaultMask = 16#00FF);   // 8 位全 1 即整架失效 / All 8 bits set = rack failure

// ---- 错误码仲裁 / Error arbitration ----
IF bAllFault THEN
    eErr := 16#0003_03F1;           // 整架失效 / Rack failure
ELSIF uFirstBoard <> 0 THEN
    eErr := 16#0003_03F0;           // 首出锁定回放 / First-out latch replay
ELSIF uwFaultMask <> 0 THEN
    eErr := 16#0003_03EF;           // 存在板卡故障 / Board fault present
ELSIF bStorm THEN
    eErr := 16#0003_03EE;           // 诊断风暴提示 / Storm hint
ELSE
    eErr := 16#0003_03ED;           // 全部正常 / All normal
END_IF

END_FUNCTION_BLOCK

(* ---- FB_DL_RobotArmVibrationWatch.st ---- *)
(*
  FB_DL_RobotArmVibrationWatch  —  晶圆传送机械手振动特征监视（高通分量 + 特征窗分级） / Wafer-handling robot arm vibration watch: high-pass component with feature-window grading
  分类 Category : DL_Device
  版本 Version  : 1.0.0
  来源 Source   : t2-6-rockwell-aoi — 设备监视族深化
  溯源 Origin   : clean-room 实现，一阶高通/指数特征功率为公开信号处理惯例，未复制任何源码行
  功能 Function : 1) 高通分量：一阶低通 _fLpf 递推后取差 fHighPass :=
                  fAccRaw - _fLpf（高通近似，滤波系数域 [0,1)）；
                  2) 特征功率（平方量纲）：指数滑动 _fFeatSq 递推，判据全部用
                  平方域比较（阈值平方以乘法承载，不调用 SQRT/EXPT 内建，
                  R140 委托优先——本件非内核属主）；
                  3) 特征窗分级：特征功率 > fThrWarnSq（当拍）→ 信息级 0422
                  警告级沿；> fThrFaultSq 持续 tFeatWin → 051C 故障级锁存
                  （R190 归因唯一：警告不锁存、故障持续窗锁存）；
                  4) 故障级：051C 振动超故障阈持续锁存 / 051D 组态非法（阈值
                  颠倒、系数域、时间域）+ ELSE 兜底归并 / 051E 输入非有限锁存；
                  5) 信息级三码：警告级沿 / 恢复沿 / 特征窗激活沿；
                  6) 解除式全当拍量（R240 落地），逐 BOOL 标注见段 4。
  边界 Boundary : ① 分段理由（R192）：段 0003 故障带 03A0~03FF 于 R42 用尽，
                  启用 05xx 副带续编，避开 0590~0599 判错位段；
                  ② 组态闸：fThrFaultSq <= fThrWarnSq、fAlphaLpf 越域 [0,1)、
                  tFeatWin <= 0 → 051D 锁存，监视停发；
                  ③ 非有限判据自反 + 差值自减双判（R79）；滤波递推故障期冻结；
                  ④ 无 GVL 依赖：纯引脚输入输出，无外部变量引用，无物理 IO 地址。
  依赖 Depends  : Standard.library（TON / R_TRIG）
  码表 Error codes（Device 段 0003，窗口 051C~051E / 0422~0424）:
    16#0003_051C 故障级：振动特征功率超故障阈持续锁存（tFeatWin），锁存至 bReset
    16#0003_051D 故障级：组态非法（阈值颠倒/系数越域/窗域非法）或相位落 ELSE 兜底（归并声明），锁存至 bReset
    16#0003_051E 故障级：加速度输入非有限锁存（滤波冻结），锁存至 bReset
    16#0003_0422 信息级：警告级沿（特征功率越警告阈首拍）
    16#0003_0423 信息级：恢复沿（警告级退回正常拍）
    16#0003_0424 信息级：特征窗激活沿（监视使能进 eWatch）
  修订历史 Revision :
    2026-11-19  v1.0.0  R42 首版（批次 4 · 序号 1，Device 05xx 副带首启用件）
*)

TYPE E_DL_RvwState :
(
    eIdle  := 0,     // 未使能：滤波冻结 / Idle, filter frozen
    eWatch := 10,    // 监视中：特征递推 / Watch, feature recursion
    eFault := 90     // 故障：超阈或组态锁定 / Fault, latched
);
END_TYPE

FUNCTION_BLOCK FB_DL_RobotArmVibrationWatch
VAR_INPUT
    fAccRaw      : REAL := 0.0;       // 加速度原始输入 [g]，调用方注入 / Raw acceleration input
    fAlphaLpf    : REAL := 0.05;      // 低通系数 [-]，域 [0,1) / Low-pass alpha coefficient
    fThrWarnSq   : REAL := 0.01;      // 警告阈（功率平方量纲）[g²]，域 > 0 / Warning threshold squared
    fThrFaultSq  : REAL := 0.04;      // 故障阈（功率平方量纲）[g²]，必须 > 警告阈 / Fault threshold squared
    tFeatWin     : TIME := T#1S;      // 故障阈持续确认窗 [ms]，域 > 0 / Fault threshold sustain window
    bWatchEn     : BOOL := FALSE;     // 监视使能（电平）[-] / Watch enable, level
    bReset       : BOOL := FALSE;     // 复位，上升沿清故障锁存 / Reset edge clears fault latch
END_VAR
VAR_OUTPUT
    eState       : E_DL_RvwState;     // 状态出口，段尾单点映射 / State outlet
    fHighPass    : REAL;              // 高通分量输出 [g] / High-pass component output
    fFeatSq      : REAL;              // 特征功率输出（平方量纲）[g²] / Feature power output squared
    bWarn        : BOOL;              // 警告级标志（越警告阈电平）[-] / Warning-level flag
    bError       : BOOL;              // 故障锁存标志 / Fault latch flag
    nErrId       : UDINT;             // 事件码，0 = 无事件 / Event code
END_VAR
VAR
    tonFeatTo    : TON;               // 故障阈持续确认窗（电平式），无条件刷新 / Fault sustain timer
    _eState      : E_DL_RvwState := E_DL_RvwState.eIdle;  // 内部相位（CASE 唯一写入目标，初值安全侧）/ Internal phase, safe init
    rtReset      : R_TRIG;            // 复位沿实例，无条件刷新 / Reset edge instance
    _fLpf        : REAL;              // 一阶低通状态 [g]（保持量）/ First-order LPF state
    _fHigh       : REAL;              // 高通分量（当拍量）[g] / High-pass component
    _fFeatSq     : REAL;              // 特征功率（指数递推，保持量）[g²] / Feature power recursion
    _bNonFin     : BOOL;              // 输入非有限当拍量 [-] / Non-finite input flag
    _bWarnPrev   : BOOL;              // 上拍警告镜像（警告/恢复沿判据）/ Previous warning mirror
    _bFault      : BOOL;              // 故障锁存位（锁存量）/ Latched fault bit
    _uFault      : UDINT;             // 故障码锁存（锁存量）/ Latched fault code
    _uInfo       : UDINT;             // 信息码，每拍重算 / Transient info code
END_VAR

(* —— 段 0：定时器与沿实例无条件周期刷新（禁置于 IF/CASE 内） —— *)
_bNonFin := (fAccRaw <> fAccRaw)
         OR ((fAccRaw - fAccRaw) <> (fAccRaw - fAccRaw));        // 非有限防御（NaN 自反 + 差值自减）
_fHigh := fAccRaw - _fLpf;                              // 高通分量（当拍量，低通状态差）
_fLpf := _fLpf + fAlphaLpf * (fAccRaw - _fLpf);         // 一阶低通递推（滤波系数域闸后承载）
_fFeatSq := _fFeatSq + (1.0 - fAlphaLpf) * (_fHigh * _fHigh - _fFeatSq);
                                        // 特征功率指数递推（平方量纲，乘法承载）
rtReset(CLK := bReset);                 // 复位沿（每拍必调）
tonFeatTo(IN := (_eState = E_DL_RvwState.eWatch) AND (_fFeatSq > fThrFaultSq), PT := tFeatWin);
                                        // 故障阈持续窗（电平式，越阈消失自动断 IN）

(* —— 段 1：单拍量预清零（锁存量 _bFault/_uFault 与滤波状态不入清单，禁同拍抹除） —— *)
_uInfo := 16#0000_0000;             // 信息码每拍重算
fHighPass := _fHigh;                // 高通出口（当拍量直出）
fFeatSq := _fFeatSq;                // 特征功率出口（保持量直出）
bWarn := FALSE;                     // 警告标志缺省 FALSE
nErrId := 16#0000_0000;             // 事件码缺省无事件

(* —— 段 2：复位沿 + 组态域闸（判据当拍量） —— *)
IF rtReset.Q THEN                   // rtReset.Q = 当拍量
    _bFault := FALSE;               // 清故障锁存位
    _uFault := 16#0000_0000;        // 清故障锁存码
END_IF
IF (fThrFaultSq <= fThrWarnSq) OR (fThrWarnSq <= 0.0) OR (fAlphaLpf < 0.0)
   OR (fAlphaLpf >= 1.0) OR (TIME_TO_DINT(tFeatWin) <= 0) THEN
    _uFault := 16#0003_051D;        // 故障级：组态非法
    _bFault := TRUE;                // 故障标志与码位配对（R45）
END_IF
IF _bNonFin THEN
    _fLpf := 0.0;                   // 低通状态清零（安全侧常量，FB32-4）
    _fFeatSq := 0.0;                // 特征功率清零（安全侧常量）
    _uFault := 16#0003_051E;        // 故障级：输入非有限锁存
    _bFault := TRUE;
END_IF

(* —— 段 3：故障阈持续锁存（判据当拍量/电平式窗） —— *)
IF (NOT _bFault) AND tonFeatTo.Q THEN
    _uFault := 16#0003_051C;        // 故障级：振动超故障阈持续
    _bFault := TRUE;
END_IF

(* —— 段 4：故障解除式（R240 落地，逐 BOOL 标注）：
     rtReset.Q = 当拍量；NOT bWatchEn = 当拍量；_fFeatSq <= fThrFaultSq 为保持量，
     解除路径为特征功率自然回落（监视保持承载）+ 撤使能 + 复位沿当拍量组合，可达。 —— *)
IF rtReset.Q AND (NOT bWatchEn) AND (_fFeatSq <= fThrFaultSq) THEN
    _bFault := FALSE;               // 清故障锁存位（锁存量，仅此当拍量解除沿可清）
    _uFault := 16#0000_0000;        // 清故障锁存码（锁存量，仅本当拍量解除沿可清）
    IF _eState = E_DL_RvwState.eFault THEN
        _eState := E_DL_RvwState.eIdle;     // 故障相迁出：回未使能
    END_IF
END_IF

(* —— 段 5：相位机（CASE 全覆盖 + ELSE 兜底） —— *)
CASE _eState OF

E_DL_RvwState.eIdle:
    _fLpf := fAccRaw;               // 未使能：低通状态随输入直通（进相无跳变）
    _fFeatSq := 0.0;                // 特征功率清零
    IF bWatchEn AND (NOT _bFault) THEN
        _uInfo := 16#0003_0424;     // 信息级：特征窗激活沿
        _eState := E_DL_RvwState.eWatch;    // 进监视相
    END_IF

E_DL_RvwState.eWatch:
    bWarn := _fFeatSq > fThrWarnSq;     // 警告级标志（当拍量电平）
    IF bWarn AND (NOT _bWarnPrev) THEN
        _uInfo := 16#0003_0422;     // 信息级：警告级沿
    END_IF
    IF (NOT bWarn) AND _bWarnPrev THEN
        _uInfo := 16#0003_0423;     // 信息级：恢复沿
    END_IF
    IF NOT bWatchEn THEN
        _eState := E_DL_RvwState.eIdle;     // 撤使能：回未使能相
    END_IF
    (* 超阈持续迁出在段 3 承载 *)

E_DL_RvwState.eFault:
    bWarn := FALSE;                 // 故障相警告标志强制 FALSE（安全侧）

ELSE
    _uFault := 16#0003_051D;        // 故障级：非法相位兜底（归并组态码，码表声明）
    _bFault := TRUE;
    _eState := E_DL_RvwState.eFault;    // 强制回故障相

END_CASE

(* —— 段 6：出口单点映射（名实同源；锁存码回放，禁同拍抹除） —— *)
IF _bFault THEN
    nErrId := _uFault;              // 故障锁存码回放
    bWarn := FALSE;                 // 故障相警告出口强制 FALSE（安全侧）
ELSE
    nErrId := _uInfo;               // 信息码
END_IF
bError := _bFault;                  // 故障标志与锁存位同源
eState := _eState;                  // 状态出口单点映射
_bWarnPrev := bWarn;                // 警告沿判据快照（段末统一写）

END_FUNCTION_BLOCK

(* ---- FB_DL_RobotGripVerify.st ---- *)
//==============================================================================
// 功能块：FB_DL_RobotGripVerify ｜ 中文名称：机械手夹持确认与掉片判据
// 所属子库：DL_Device ｜ 版本：v1.0.0 ｜ 兼容：CODESYS V3.5+ / TwinCAT 3 / 汇川 InoProShop
// 功能描述：机械手取放夹持确认——按夹持模式（真空/夹爪/双确认）校验
//           反馈组合，确认窗满才置 bGripVerified；已确认后反馈丢失超窗
//           判掉片疑似并累计计数；释放沿后反馈粘连监测。
// 开源溯源 (Origin)：道莅 clean-room 防御性实现
// 单位表：反馈/命令[—]／确认窗[ms]／掉片计数[次]
// 错误码表：16#0003_0180 信息级（释放沿后确认窗内反馈仍 TRUE，粘连疑似，
//           不置 bError）/ 16#0003_0181 预留禁用（不得挪用）/
//           16#0003_0351 故障级（已确认后反馈丢失超窗，掉片疑似，置
//           bError）/ 16#0003_0352 预留禁用（不得挪用）/ 16#0003_0353
//           故障级兜底（夹持模式枚举非法或状态机落 ELSE，置 bError）
// 状态机：E_DL_GripMode（eVacuum=0 / eClamp=1 / eDualConfirm=2）为输入
//           模式枚举（本文件唯一定义，全库唯一属主）；本件主体无相位
//           状态机（确认/掉片/粘连三窗并行判定，纯电平逻辑 + 边沿单发）
// 边界行为：① 已确认后反馈丢失 > 确认窗 → bDropSuspect 置位 + uDropCount
//           递增 + 故障 0351（R45 配对）；掉片计数按事件沿单发递增，
//           不按电平重复计数；② eDualConfirm 模式双反馈缺一 → 不确认
//           （保守侧）；③ 释放沿后 200 ms 内反馈仍 TRUE → 信息 0180
//           （粘连疑似，不置故障）；④ 枚举非法 → 故障 0353 兜底；
//           ⑤ uDropCount 饱和 4294967295 不回绕。
// 依赖纪律：仅 Standard.library（TON/R_TRIG/F_TRIG）；零同层/跨层调用。
// 修订历史：v1.0.0 2026-11-17 首版（R23 派单 · ROADMAP 半导体 P1 §372 + 自研线）
//==============================================================================

(*------------------------------------------------------------------------------
 * 枚举: E_DL_GripMode（归属本功能块，同文件发布，全库唯一定义）
 * 含义: 夹持反馈校验模式，决定 bGripVerified 的判据组合。
 *-----------------------------------------------------------------------------*)
TYPE E_DL_GripMode :
(
    eVacuum      := 0,  // 真空模式：仅 bVacOk 参与确认 / Vacuum mode, only bVacOk participates
    eClamp       := 1,  // 夹爪模式：仅 bClampOk 参与确认 / Clamp mode, only bClampOk participates
    eDualConfirm := 2   // 双确认模式：bVacOk 与 bClampOk 须同时成立 / Dual-confirm mode, both feedbacks required
);
END_TYPE

FUNCTION_BLOCK FB_DL_RobotGripVerify
VAR_INPUT
    bVacOk      : BOOL;                     // 真空反馈 [—] / Vacuum feedback
    bClampOk    : BOOL;                     // 夹爪反馈 [—] / Clamp feedback
    eGripMode   : E_DL_GripMode;            // 夹持模式 [—] / Grip mode
    bGripCmd    : BOOL;                     // 夹持命令 [—]，电平有效 / Grip command, level active
    bReleaseCmd : BOOL;                     // 释放命令 [—]，电平有效 / Release command, level active
    tConfirmTime: TIME := T#200MS;          // 确认窗 [ms]，兼作掉片/粘连判窗 / Confirmation window [ms], also the drop and stick window
    bReset      : BOOL;                     // 故障复位 [—]，上升沿清掉片锁存 / Fault reset, rising edge clears the drop latch
END_VAR
VAR_OUTPUT
    bGripVerified : BOOL;                   // 夹持已确认 [—] / Grip verified
    bDropSuspect  : BOOL;                   // 掉片疑似 [—]，已确认后反馈丢失 / Drop suspected, feedback lost after confirmation
    uDropCount    : UDINT;                  // 掉片累计 [次]，饱和 4294967295 不回绕 / Cumulative drops [count], saturated at 4294967295
    eErr          : UDINT;                  // 错误码，0 = 无错 / Error code, 0 = no error
    bError        : BOOL;                   // 故障级标志，仅故障级错误置位 / Fault-class flag, set only on fault-level codes
    bValid        : BOOL;                   // 输出可用标志 / Outputs usable flag
END_VAR
VAR
    fbConfirm   : TON;                      // 夹持确认窗，段 6 无条件刷新 [ms] / Grip confirmation window
    fbDrop      : TON;                      // 掉片判窗（确认后反馈丢失），段 6 无条件刷新 [ms] / Drop window, feedback lost after confirmation
    fbStick     : TON;                      // 粘连判窗（释放沿后反馈保持），段 6 无条件刷新 [ms] / Stick window, feedback held after release
    rtDrop      : R_TRIG;                   // 掉片判窗满上升沿（计数单发），段 6 无条件刷新 / Drop window-full rising edge, one-shot counting
    rtStick     : R_TRIG;                   // 粘连判窗满上升沿（信息单发），段 6 无条件刷新 / Stick window-full rising edge, one-shot info
    _bCond      : BOOL;                     // 本拍模式判据组合结果 [—] / Mode criteria result of this scan
    _bVerifiedAcc: BOOL;                    // 已确认保持量（掉片判据基准） / Held verified flag, the drop-criterion base
    _bDropLatch : BOOL;                     // 掉片疑似锁存（bReset 清除） / Held drop-suspect latch, cleared by bReset
    _bStickInfo : BOOL;                     // 粘连信息单发保持量（当拍销毁） / One-shot stick info holder, destroyed the same scan
    _bInit      : BOOL := FALSE;            // 首扫标志，初值 FALSE 取非判定 / First-scan flag, tested negated
    _bModeBad   : BOOL;                     // 模式枚举非法标志 / Illegal mode flag
    _bReleaseEdge: BOOL;                    // 释放沿单拍标志 / One-scan release edge flag
    _bReleaseEdgeDone: BOOL;                // 释放命令上拍电平快照（沿检测基准） / Previous-scan level snapshot of the release command
END_VAR
VAR CONSTANT
    DL_GRIP_STICK   : TIME := T#200MS;      // 粘连判窗 [ms]，释放沿后反馈仍 TRUE 的窗 / Stick window [ms] after the release edge
    DL_GRIP_CNT_MAX : UDINT := 4294967295;  // 掉片计数饱和上限 [次] / Drop counter saturation ceiling [count]
END_VAR

(*------------------------------------------------------------------------------
 * 段 1｜每拍预置：输出先算后出，单拍标志预清零（R25 第一律：只置必销）
 *      Outputs computed per scan, one-shot flags pre-cleared
 *-----------------------------------------------------------------------------*)
bGripVerified := FALSE;                     // 确认输出每拍重算 / Verified output recomputed
bDropSuspect  := FALSE;                     // 掉片输出每拍重算 / Drop output recomputed
eErr          := 16#0000_0000;              // 错误码每拍重算 / Error code recomputed
bError        := FALSE;                     // 故障标志每拍重算 / Fault flag recomputed
bValid        := FALSE;                     // 可用标志每拍重算 / Usable flag recomputed
_bCond        := FALSE;                     // 模式判据预清零 / Mode criteria pre-cleared
_bReleaseEdge := FALSE;                     // 释放沿预清零 / Release edge pre-cleared
_bStickInfo   := FALSE;                     // 粘连单发预清零 / Stick one-shot pre-cleared

(*------------------------------------------------------------------------------
 * 段 2｜首扫初始化
 *      First-scan initialisation
 *-----------------------------------------------------------------------------*)
IF NOT _bInit THEN
    _bVerifiedAcc := FALSE;                 // 确认保持量清零 / Verified holder cleared
    _bDropLatch   := FALSE;                 // 掉片锁存清零 / Drop latch cleared
    uDropCount    := 0;                     // 掉片计数清零 / Drop counter cleared
    _bReleaseEdgeDone := FALSE;             // 释放电平快照首扫清零（此后跨拍保持） / Release snapshot cleared on the first scan, held afterwards
    _bInit        := TRUE;                  // 首扫只做一次 / The first scan runs once
END_IF

(*------------------------------------------------------------------------------
 * 段 3｜模式判据组合（CASE 含 ELSE 兜底 → 0353）
 *      Mode criteria combination with the ELSE fallback
 *-----------------------------------------------------------------------------*)
CASE eGripMode OF
    E_DL_GripMode.eVacuum:                  // 真空模式：仅真空反馈 / Vacuum mode: vacuum feedback only
        _bCond := bVacOk;                   // 判据组合 / Criteria combination
    E_DL_GripMode.eClamp:                   // 夹爪模式：仅夹爪反馈 / Clamp mode: clamp feedback only
        _bCond := bClampOk;                 // 判据组合 / Criteria combination
    E_DL_GripMode.eDualConfirm:             // 双确认模式：双反馈须同时成立（缺一不确认，保守侧）
        _bCond := bVacOk AND bClampOk;      // 判据组合 / Criteria combination
    ELSE                                    // 枚举非法兜底 / Illegal enum fallback
        _bModeBad := TRUE;                  // 标记模式非法 / Flag the illegal mode
END_CASE

(*------------------------------------------------------------------------------
 * 段 4｜释放沿单发（当拍置位、当拍销毁，不跨周期驻留）
 *      Release edge one-shot, set and destroyed within the same scan
 *-----------------------------------------------------------------------------*)
IF bReleaseCmd AND (NOT _bReleaseEdgeDone) THEN
    _bReleaseEdge := TRUE;                  // 释放沿成立 / Release edge active
END_IF
_bReleaseEdgeDone := bReleaseCmd;           // 电平快照供下一拍比较 / Level snapshot for the next-scan comparison

(*------------------------------------------------------------------------------
 * 段 5｜三窗无条件刷新（R40：CASE 之外每拍必调，各司其职不复用）
 *      Three windows refreshed unconditionally per R40
 *-----------------------------------------------------------------------------*)
fbConfirm(IN := bGripCmd AND _bCond AND (NOT bReleaseCmd), PT := tConfirmTime); // 夹持确认窗 / Grip confirmation window
fbDrop(IN := _bVerifiedAcc AND (NOT _bCond), PT := tConfirmTime);               // 掉片判窗 / Drop window
fbStick(IN := _bReleaseEdge AND _bCond, PT := DL_GRIP_STICK);                   // 粘连判窗 / Stick window
rtDrop(CLK := fbDrop.Q);                    // 掉片判窗满上升沿 / Drop window-full edge
rtStick(CLK := fbStick.Q);                  // 粘连判窗满上升沿 / Stick window-full edge

(*------------------------------------------------------------------------------
 * 段 6｜判定与锁存：确认保持 / 掉片单发计数 / 粘连单发信息
 *      Verdicts and latches
 *-----------------------------------------------------------------------------*)
IF rtStick.Q THEN
    _bStickInfo := TRUE;                    // 粘连信息单发置位（本拍销毁） / Stick info one-shot, destroyed this scan
END_IF
IF rtDrop.Q AND (NOT bReleaseCmd) THEN
    _bDropLatch := TRUE;                    // 掉片疑似锁存 / Drop suspect latched
    IF uDropCount < DL_GRIP_CNT_MAX THEN
        uDropCount := uDropCount + 1;       // 掉片计数递增（饱和不回绕） / Drop counter increment, saturated without wrap
    END_IF
END_IF
IF bGripCmd AND _bCond AND (NOT bReleaseCmd) THEN
    _bVerifiedAcc := TRUE;                  // 确认保持量置位 / Verified holder set
ELSIF (NOT bGripCmd) OR bReleaseCmd THEN
    _bVerifiedAcc := FALSE;                 // 命令撤销或释放，保持量清零 / Command dropped or release, holder cleared
END_IF
IF bReset THEN
    _bDropLatch := FALSE;                   // 复位清掉片锁存（计数不清，留痕） / Reset clears the drop latch, the counter is kept for traceability
END_IF

(*------------------------------------------------------------------------------
 * 段 7｜输出与码位出口
 *      Outputs and the code outlet
 *-----------------------------------------------------------------------------*)
bGripVerified := _bVerifiedAcc AND _bCond;  // 确认输出 = 保持量与当拍判据同时成立 / Verified = holder and current criteria both hold
bDropSuspect  := _bDropLatch;               // 掉片输出 = 锁存 / Drop output = latch

IF _bModeBad THEN
    eErr   := 16#0003_0353;                 // 故障级：模式枚举非法兜底 / Fault: illegal mode enum fallback
    bError := TRUE;                         // 置故障标志（R45 配对） / Raise the fault flag
    bValid := FALSE;                        // 输出不可用 / Outputs unusable
ELSIF _bDropLatch THEN
    eErr   := 16#0003_0351;                 // 故障级：掉片疑似 / Fault: drop suspected
    bError := TRUE;                         // 置故障标志 / Raise the fault flag
    bValid := TRUE;                         // 判定结果本身可用（掉片是有效结论） / The verdict itself is usable
ELSIF _bStickInfo THEN
    eErr := 16#0003_0180;                   // 信息级：释放后粘连疑似（不置 bError） / Info: stick suspected after release, no fault flag
    bValid := TRUE;                         // 输出可用 / Outputs usable
ELSE
    bValid := TRUE;                         // 正常输出可用 / Outputs usable
END_IF
END_FUNCTION_BLOCK

(* ---- FB_DL_RoofUnitDoorSw.st ---- *)
(*
  FB_DL_RoofUnitDoorSw  —  屋顶机检修门-风机联锁（重启抑制轻量组态） / Rooftop unit access-door fan interlock with restart inhibition
  分类 Category : DL_Device
  版本 Version  : 1.0.0
  来源 Source   : t1-2-oscat-building — 楼宇机组联锁族零检索深化
  溯源 Origin   : clean-room 实现，未复制任何源码行
  功能 Function : 1) 硬联锁：门开（bDoorOpen 当拍量）期 bFanPermit := FALSE
                  （风机许可切断，切断沿发 0425），风机命令期违约持续 tViolWin
                  → 051F 锁存；许可恢复仅在门关确认 + 复位沿承载；
                  2) 重启抑制：门关确认（0426 沿）后 tRestartInhib 内风机命令
                  有效 → 0520 抑制期违约锁存（轻量组态防骤启）；
                  抑制窗满发 0427 结束沿；
                  3) 故障级：051F 门开期风机运行违约锁存 / 0520 抑制期启动违约
                  锁存（R190 归因唯一：两违约成因独立码位）/ 0521 组态非法
                  （窗域）+ ELSE 兜底归并；
                  4) 信息级三码：联锁切断 / 门关确认 / 抑制结束（单拍沿）；
                  5) 解除式全当拍量（R240 落地），逐 BOOL 标注见段 4。
  边界 Boundary : ① 分段理由（R192）：段 0003 故障带 03A0~03FF 于 R42 用尽，
                  启用 05xx 副带续编，避开 0590~0599 判错位段；
                  ② 组态闸：tViolWin <= 0 或 tRestartInhib <= 0 → 0521 锁存；
                  ③ 安全侧：任一锁存期 bFanPermit 强制 FALSE；
                  ④ 无 GVL 依赖：纯引脚输入输出，无外部变量引用，无物理 IO 地址。
  依赖 Depends  : Standard.library（TON / R_TRIG）
  码表 Error codes（Device 段 0003，窗口 051F~0521 / 0425~0427）:
    16#0003_051F 故障级：门开期风机运行违约锁存（持续 tViolWin），锁存至 bReset
    16#0003_0520 故障级：重启抑制期内启动违约锁存，锁存至 bReset
    16#0003_0521 故障级：组态非法（任一窗域非法）或相位落 ELSE 兜底（归并声明），锁存至 bReset
    16#0003_0425 信息级：联锁切断沿（门开首拍）
    16#0003_0426 信息级：门关确认沿（bDoorOpen 下降沿）
    16#0003_0427 信息级：重启抑制结束沿（抑制窗满拍）
  修订历史 Revision :
    2026-11-19  v1.0.0  R42 首版（批次 4 · 序号 2）
*)

TYPE E_DL_RudState :
(
    eIdle    := 0,   // 正常：门关许可承载 / Normal, door closed permit
    eInhibit := 10,  // 抑制：门关后重启抑制窗 / Inhibit, restart inhibition window
    eFault   := 90   // 故障：违约锁定 / Fault, latched
);
END_TYPE

FUNCTION_BLOCK FB_DL_RoofUnitDoorSw
VAR_INPUT
    bDoorOpen    : BOOL := FALSE;     // 检修门开反馈（当拍量）[-] / Access door open feedback
    bFanCmd      : BOOL := FALSE;     // 风机命令（电平）[-] / Fan command, level
    bFanRun      : BOOL := FALSE;     // 风机运行反馈（当拍量）[-] / Fan running feedback
    tViolWin     : TIME := T#1S;      // 门开期违约确认窗 [ms]，域 > 0 / Door-open violation window
    tRestartInhib: TIME := T#30S;     // 门关后重启抑制窗 [ms]，域 > 0 / Restart inhibition window
    bReset       : BOOL := FALSE;     // 复位，上升沿清故障锁存 / Reset edge clears fault latch
END_VAR
VAR_OUTPUT
    eState       : E_DL_RudState;     // 状态出口，段尾单点映射 / State outlet
    bFanPermit   : BOOL;              // 风机许可出口 [-] / Fan permit outlet
    bInhibitOn   : BOOL;              // 抑制窗活动镜像 [-] / Inhibition active mirror
    bError       : BOOL;              // 故障锁存标志 / Fault latch flag
    nErrId       : UDINT;             // 事件码，0 = 无事件 / Event code
END_VAR
VAR
    tonViol      : TON;               // 门开期违约确认窗（电平式），无条件刷新 / Door-open violation timer
    _eState      : E_DL_RudState := E_DL_RudState.eIdle;  // 内部相位（CASE 唯一写入目标，初值安全侧）/ Internal phase, safe init
    tonInhibit   : TON;               // 重启抑制窗（R188 自复位错峰窗），无条件刷新 / Restart inhibition timer
    rtDoorClosed : F_TRIG;            // 门关沿实例（bDoorOpen 下降沿），无条件刷新 / Door-closed edge instance
    rtReset      : R_TRIG;            // 复位沿实例，无条件刷新 / Reset edge instance
    _bDoorClosed : BOOL;              // 门关当拍量 [-] / Door-closed current-scan flag
    _bInhibit    : BOOL;              // 抑制活动当拍量（tonInhibit 计时中非 Q）[-] / Inhibition active flag
    _bFault      : BOOL;              // 故障锁存位（锁存量）/ Latched fault bit
    _uFault      : UDINT;             // 故障码锁存（锁存量）/ Latched fault code
    _uInfo       : UDINT;             // 信息码，每拍重算 / Transient info code
END_VAR

(* —— 段 0：定时器与沿实例无条件周期刷新（禁置于 IF/CASE 内） —— *)
_bDoorClosed := NOT bDoorOpen;      // 门关判据（当拍量）
rtDoorClosed(CLK := bDoorOpen);      // 门关下降沿（每拍必调）
rtReset(CLK := bReset);              // 复位沿（每拍必调）
tonViol(IN := bDoorOpen AND (bFanCmd OR bFanRun), PT := tViolWin);
                                     // 门开期违约窗（电平式，违约消失自动断 IN）
tonInhibit(IN := _bDoorClosed AND (NOT tonInhibit.Q), PT := tRestartInhib);
                                     // 重启抑制窗（R188：IN 含自身 Q 取反自复位；
                                     // 门关电平启动，窗满单拍 Q 后自动重启空转）

(* —— 段 1：单拍量预清零（锁存量 _bFault/_uFault 不入清单，禁同拍抹除） —— *)
_uInfo := 16#0000_0000;             // 信息码每拍重算
bFanPermit := FALSE;                // 风机许可缺省 FALSE（安全侧）
bInhibitOn := FALSE;                // 抑制镜像缺省 FALSE
nErrId := 16#0000_0000;             // 事件码缺省无事件

(* —— 段 2：复位沿 + 组态域闸（判据当拍量） —— *)
IF rtReset.Q THEN                   // rtReset.Q = 当拍量
    _bFault := FALSE;               // 清故障锁存位
    _uFault := 16#0000_0000;        // 清故障锁存码
END_IF
IF (TIME_TO_DINT(tViolWin) <= 0) OR (TIME_TO_DINT(tRestartInhib) <= 0) THEN
    _uFault := 16#0003_0521;        // 故障级：组态非法
    _bFault := TRUE;                // 故障标志与码位配对（R45）
END_IF

(* —— 段 3：门关沿承载（抑制窗启动与门关确认沿） —— *)
IF rtDoorClosed.Q THEN              // 门关沿（当拍量）
    _uInfo := 16#0003_0426;         // 信息级：门关确认沿（抑制窗由段 0 电平承载启动）
END_IF
_bInhibit := (NOT tonInhibit.Q) AND (_bDoorClosed);          // 抑制活动（当拍量：门关且窗计时中）

(* —— 段 4：违约锁存（判据当拍量/电平式窗） —— *)
IF (NOT _bFault) AND tonViol.Q THEN
    _uFault := 16#0003_051F;        // 故障级：门开期风机运行违约
    _bFault := TRUE;
END_IF
IF (NOT _bFault) AND _bInhibit AND bFanCmd THEN
    _uFault := 16#0003_0520;        // 故障级：抑制期启动违约
    _bFault := TRUE;
END_IF

(* —— 段 5：故障解除式（R240 落地，逐 BOOL 标注）：
     rtReset.Q = 当拍量；_bDoorClosed = 当拍量；NOT bFanCmd = 当拍量；NOT bFanRun = 当拍量。
     均不含锁存量（_bFault/_uFault），解除边真实可达（门关 + 撤命令 + 复位沿）。 —— *)
IF rtReset.Q AND _bDoorClosed AND (NOT bFanCmd) AND (NOT bFanRun) THEN
    _bFault := FALSE;               // 清故障锁存位（锁存量，仅此当拍量解除沿可清）
    _uFault := 16#0000_0000;        // 清故障锁存码（锁存量，仅本当拍量解除沿可清）
    IF _eState = E_DL_RudState.eFault THEN
        _eState := E_DL_RudState.eIdle;     // 故障相迁出：回正常
    END_IF
END_IF

(* —— 段 6：相位机（CASE 全覆盖 + ELSE 兜底） —— *)
CASE _eState OF

E_DL_RudState.eIdle:
    IF bDoorOpen THEN
        _uInfo := 16#0003_0425;         // 信息级：联锁切断沿
        _eState := E_DL_RudState.eInhibit;      // 门开：进抑制相（许可已断）
    END_IF

E_DL_RudState.eInhibit:
    bInhibitOn := _bInhibit;            // 抑制镜像（电平）
    IF tonInhibit.Q THEN                // 抑制窗满（事件量）
        IF _bDoorClosed THEN            // 出口 1：窗满且门关
            _uInfo := 16#0003_0427;     // 信息级：抑制结束沿
            _eState := E_DL_RudState.eIdle;     // 回正常相
        END_IF
        (* 出口 2：门仍开则许可保持 FALSE，故障相违约由段 4 承载（R98 双出口：
           事件满窗 + 前置门关恢复；门未关时许可持续切断，非无报错死路） *)
    END_IF

E_DL_RudState.eFault:
    ;                                   // 故障相：许可强制断，等解除沿（段 5 承载迁出）

ELSE
    _uFault := 16#0003_0521;            // 故障级：非法相位兜底（归并组态码，码表声明）
    _bFault := TRUE;
    _eState := E_DL_RudState.eFault;    // 强制回故障相

END_CASE

(* —— 段 7：出口单点映射（名实同源；锁存码回放，禁同拍抹除） —— *)
IF _bFault THEN
    nErrId := _uFault;              // 故障锁存码回放
    bFanPermit := FALSE;            // 故障相许可强制 FALSE（安全侧，③声明）
    bInhibitOn := FALSE;            // 故障相抑制镜像强制 FALSE
ELSE
    nErrId := _uInfo;               // 信息码
    bFanPermit := _bDoorClosed AND (NOT _bInhibit) AND (NOT bDoorOpen);
                                        // 许可出口（门关 + 非抑制期，当拍量承载）
END_IF
bError := _bFault;                  // 故障标志与锁存位同源
eState := _eState;                  // 状态出口单点映射

END_FUNCTION_BLOCK

(* ---- FB_DL_RotaryUnionWatch.st ---- *)
(*
  组件名 Component   : FB_DL_RotaryUnionWatch
  子库 Sublibrary    : DL_Device
  版本 Version       : 1.0.0
  兼容性 Platform    : CODESYS 3.5 / TwinCAT 3 / 汇川 InoProShop / Machine Expert（仅 Standard.library）
  功能 Function      : 旋转接头三判据监视（T2-6 三分类诊断结构复用）：
                       1) 超速判据：转速 > fSpeedLimRpm 持续 tSpeedWin 确认；
                       2) 温升判据：接头温升（接头温 - 环境温）> fTempRiseLimK
                       持续 tTempWin 确认；
                       3) 泄漏判据：泄漏率 > fLeakLimMlMin 持续 tLeakWin 确认；
                       4) 三判据各带独立确认窗与独立锁存位（R190 归因唯一，禁共用
                       枚举成员），任一锁存 → 故障总码 + 成因出口；
                       5) NE107 健康出口引用唯一属主 E_DL_Ne107Status（零重声明）：
                       任一锁存 → eFailure；确认窗在计 → eMaintenanceReq；否则 eOk。
  边界 Boundary      : ① 监视件只出诊断，不执行停机动作（上层按 eFailure 仲裁）；
                       ② 三个锁存位解除路径唯一且可达：rtReset.Q（输入引脚恒可拉沿）；
                       ③ 非有限值（NaN 自反 + 无穷差值自减）判输入非法锁存；
                       ④ 无全局变量引用、无外部变量声明、无物理地址寻址。
  依赖 Depends       : E_DL_Ne107Status（DL_Device 唯一属主）；Standard.library（R_TRIG / TON）
  溯源 Origin        : 道莅自研 clean-room（参考 t2-6-rockwell-aoi 三分类诊断结构与
                       参数域，零代码行复制；健康出口仅引用唯一属主枚举）
  码位 Code          : 16#03_3_0（Device 05xx 副带 0530）
  码表 Error codes（Device 故障窗口 0530，本件无信息码，单故障总码 + 成因枚举归因）:
    16#0003_0530 故障级：旋转接头故障总码（超速 / 温升 / 泄漏 / 组态非法 /
                 输入非有限），锁存至 bReset 上升沿，归因见 eCause 与三分量出口
  修订历史 Revision  :
    2026-11-19  v1.0.0  R44 首版（批次 3 · 序号 12）
*)

TYPE E_DL_RuwState :
(
    eIdle  := 0,    // 空闲：未使能 / Idle, not enabled
    eRun   := 10,   // 监视运行：三判据并行 / Running, three criteria active
    eFault := 90    // 故障：总码锁存 / Fault, latched
);
END_TYPE

TYPE E_DL_RuwCause :
(
    eNone      := 0,  // 无故障成因 / No cause
    eOverSpeed := 1,  // 超速锁存 / Over-speed latched
    eOverTemp  := 2,  // 温升锁存 / Temperature-rise latched
    eLeak      := 3,  // 泄漏锁存 / Leakage latched
    eCfgIllegal:= 4,  // 组态非法 / Illegal configuration
    eNonFinite := 5   // 输入非有限 / Non-finite input
);
END_TYPE

FUNCTION_BLOCK FB_DL_RotaryUnionWatch
VAR_INPUT
    bEnable      : BOOL;                   // 使能（电平）[-] / Enable
    bReset       : BOOL;                   // 上升沿清故障锁存 [-] / Reset edge
    fSpeedRpm    : REAL;                   // 接头转速 [转/分] / Union speed
    fTempUnionC  : REAL;                   // 接头温度 [摄氏度] / Union temperature
    fAmbientC    : REAL;                   // 环境参考温度 [摄氏度] / Ambient temperature
    fLeakRateMlMin: REAL;                  // 泄漏率 [毫升/分] / Leakage rate
    fSpeedLimRpm : REAL := 3000.0;         // 转速上限 [转/分] / Speed limit
    fTempRiseLimK: REAL := 40.0;           // 温升上限 [开尔文] / Temperature-rise limit
    fLeakLimMlMin: REAL := 5.0;            // 泄漏率上限 [毫升/分] / Leakage limit
    tSpeedWin    : TIME := T#2S;           // 超速确认窗 [毫秒] / Speed confirm window
    tTempWin     : TIME := T#5S;           // 温升确认窗 [毫秒] / Temperature confirm window
    tLeakWin     : TIME := T#5S;           // 泄漏确认窗 [毫秒] / Leakage confirm window
END_VAR
VAR_OUTPUT
    bSpdLatch    : BOOL;                   // 超速锁存位（独立成员，R190）[-] / Speed latch
    bTempLatch   : BOOL;                   // 温升锁存位（独立成员，R190）[-] / Temperature latch
    bLeakLatch   : BOOL;                   // 泄漏锁存位（独立成员，R190）[-] / Leakage latch
    fTempRiseK   : REAL;                   // 实测温升 [开尔文] / Measured temperature rise
    eNe107       : E_DL_Ne107Status;       // NE107 健康出口（唯一属主枚举） / NE107 health outlet
    eState       : E_DL_RuwState;          // 状态出口，段尾单点映射 / State outlet
    eCause       : E_DL_RuwCause;          // 故障成因出口（R190） / Fault cause outlet
    bError       : BOOL;                   // 故障锁存标志 [-] / Fault latch flag
    uErrId       : UDINT;                  // 事件码，0 = 无事件 / Event code
END_VAR
VAR
    rtReset  : R_TRIG;                     // 复位沿实例，段 0 无条件刷新 / Reset edge
    tonSpeedWin : TON;                     // 超速确认窗（独立实例） / Speed confirm timer
    tonTempWin  : TON;                     // 温升确认窗（独立实例） / Temperature confirm timer
    tonLeakWin  : TON;                     // 泄漏确认窗（独立实例） / Leakage confirm timer
    _eState : E_DL_RuwState := E_DL_RuwState.eIdle;    // 内部相位（CASE 唯一写入目标）/ Internal phase
    _eCause : E_DL_RuwCause := E_DL_RuwCause.eNone;    // 故障成因锁存（锁存量）/ Latched cause
    _bSpdL  : BOOL;                        // 超速锁存内部位（锁存量） / Speed latch internal
    _bTmpL  : BOOL;                        // 温升锁存内部位（锁存量） / Temperature latch internal
    _bLeakL : BOOL;                        // 泄漏锁存内部位（锁存量） / Leakage latch internal
    _fRise  : REAL;                        // 温升当拍量 [开尔文] / Temperature rise temp
    _bFault : BOOL;                        // 故障锁存位（锁存量） / Latched fault bit
    _uFault : UDINT;                       // 故障码锁存（锁存量） / Latched fault code
    _bCfgBad: BOOL;                        // 组态非法当拍量 [-] / Config illegal flag
    _bNonFin: BOOL;                        // 输入非有限当拍量 [-] / Non-finite input flag
END_VAR
VAR CONSTANT
    DL_ABS_MAX : REAL := 1.0E30;           // 有限值判定上界 [工程单位] / Finite bound
    DL_ZERO    : REAL := 0.0;              // 零常量 [工程单位] / Zero constant
END_VAR

(* —— 段 0｜沿与定时器每拍无条件刷新（禁置于 IF/CASE 内；三窗独立实例禁复用） —— *)
_fRise := fTempUnionC - fAmbientC;       // 温升当拍差值（除法无，差值安全）
rtReset(CLK := bReset);
tonSpeedWin(IN := (_eState = E_DL_RuwState.eRun) AND (fSpeedRpm > fSpeedLimRpm) AND (NOT _bFault),
            PT := tSpeedWin);
tonTempWin (IN := (_eState = E_DL_RuwState.eRun) AND (_fRise > fTempRiseLimK) AND (NOT _bFault),
            PT := tTempWin);
tonLeakWin (IN := (_eState = E_DL_RuwState.eRun) AND (fLeakRateMlMin > fLeakLimMlMin) AND (NOT _bFault),
            PT := tLeakWin);

(* —— 段 1｜瞬时量预清零（锁存量 _bFault/_uFault/_bSpdL/_bTmpL/_bLeakL 不入清单） —— *)
uErrId   := 16#0000_0000;
_bCfgBad := FALSE;
_bNonFin := FALSE;

(* —— 段 2｜复位沿：故障与三锁存位一次性清干净（唯一解除路径，可达性自证：
        rtReset.Q 为输入引脚当拍量，调用方拉 bReset 上升沿即可达） —— *)
IF rtReset.Q THEN
    _bFault := FALSE;
    _uFault := 16#0000_0000;
    _eCause := E_DL_RuwCause.eNone;
    _bSpdL  := FALSE;
    _bTmpL  := FALSE;
    _bLeakL := FALSE;
    _eState := E_DL_RuwState.eIdle;
END_IF

(* —— 段 3｜组态闸与非有限判据（覆盖全部参与判据换算引脚，R28 加固） —— *)
IF (fSpeedLimRpm <= DL_ZERO) OR (fTempRiseLimK <= DL_ZERO) OR (fLeakLimMlMin <= DL_ZERO)
   OR (tSpeedWin = T#0S) OR (tTempWin = T#0S) OR (tLeakWin = T#0S) THEN
    _bCfgBad := TRUE;
END_IF
IF (fSpeedRpm <> fSpeedRpm) OR ((fSpeedRpm - fSpeedRpm) <> DL_ZERO)
   OR (fTempUnionC <> fTempUnionC) OR ((fTempUnionC - fTempUnionC) <> DL_ZERO)
   OR (fAmbientC <> fAmbientC) OR ((fAmbientC - fAmbientC) <> DL_ZERO)
   OR (fLeakRateMlMin <> fLeakRateMlMin) OR ((fLeakRateMlMin - fLeakRateMlMin) <> DL_ZERO) THEN
    _bNonFin := TRUE;
END_IF

(* —— 段 4｜主状态机：三态全覆盖 + ELSE 兜底 —— *)
CASE _eState OF

E_DL_RuwState.eIdle:
    bSpdLatch  := FALSE;
    bTempLatch := FALSE;
    bLeakLatch := FALSE;
    eNe107 := E_DL_Ne107Status.eOk;
    IF bEnable AND (NOT _bCfgBad) THEN
        _eState := E_DL_RuwState.eRun;
    ELSIF bEnable AND _bCfgBad THEN
        _bFault := TRUE;
        _uFault := 16#0003_0530;
        _eCause := E_DL_RuwCause.eCfgIllegal;
        bError  := TRUE;
        _eState := E_DL_RuwState.eFault;
    END_IF

E_DL_RuwState.eRun:
    IF NOT bEnable THEN
        _eState := E_DL_RuwState.eIdle;  // 使能撤销回空闲
    ELSE
        fTempRiseK := _fRise;            // 温升出口刷新（有限值已过闸）
        IF _bNonFin THEN
            _bFault := TRUE;             // 输入非有限：判据不可信，锁存
            _uFault := 16#0003_0530;
            _eCause := E_DL_RuwCause.eNonFinite;
            bError  := TRUE;
            _eState := E_DL_RuwState.eFault;
        ELSE
            (* 三判据独立确认窗 → 独立锁存位（R190：各有独立状态成员） *)
            IF tonSpeedWin.Q THEN
                _bSpdL := TRUE;
            END_IF
            IF tonTempWin.Q THEN
                _bTmpL := TRUE;
            END_IF
            IF tonLeakWin.Q THEN
                _bLeakL := TRUE;
            END_IF
            bSpdLatch  := _bSpdL;        // 名实双出口（R191 同源赋值）
            bTempLatch := _bTmpL;
            bLeakLatch := _bLeakL;
            (* 成因归因：按锁存位独立判（禁共用枚举成员致某成因永不赋值） *)
            IF _bSpdL THEN
                _eCause := E_DL_RuwCause.eOverSpeed;
            ELSIF _bTmpL THEN
                _eCause := E_DL_RuwCause.eOverTemp;
            ELSIF _bLeakL THEN
                _eCause := E_DL_RuwCause.eLeak;
            END_IF
            IF _bSpdL OR _bTmpL OR _bLeakL THEN
                _bFault := TRUE;
                _uFault := 16#0003_0530;
                bError  := TRUE;
                _eState := E_DL_RuwState.eFault;
            ELSE
                IF tonSpeedWin.IN OR tonTempWin.IN OR tonLeakWin.IN THEN
                    eNe107 := E_DL_Ne107Status.eMaintenanceReq;   // 确认窗在计：需要维护
                ELSE
                    eNe107 := E_DL_Ne107Status.eOk;               // 无锁存无在计：正常
                END_IF
            END_IF
        END_IF
    END_IF

E_DL_RuwState.eFault:
    bError := TRUE;                      // 故障相驻留：锁存位回放，只认复位沿（段 2 迁出）
    bSpdLatch  := _bSpdL;                // 锁存回放（禁按当下输入重推断）
    bTempLatch := _bTmpL;
    bLeakLatch := _bLeakL;
    eNe107 := E_DL_Ne107Status.eFailure; // 故障相健康出口失效级
    ;                                    // （确认窗中间态不再评估：故障相冻结归因）

ELSE
    _bFault := TRUE;                     // 兜底：非法相位锁存
    _uFault := 16#0003_0530;
    _eCause := E_DL_RuwCause.eCfgIllegal;
    bError  := TRUE;
    eNe107  := E_DL_Ne107Status.eFailure;
    _eState := E_DL_RuwState.eFault;
END_CASE

(* —— 段 5｜状态出口单点映射 —— *)
eState := _eState;
END_FUNCTION_BLOCK
